                           #diagnostics.partnerConfig.sizeOfReceiveBuffer := 0;
                           #diagnostics.partnerConfig.sizeOfSendBuffer := 0;
                           #connected := #statConnected := TRUE;
                           #statState.cfgSender := #OPERATION;

                           #statDiag.bufferIndex := #statDiag.bufferIndex + 1;
                           #statDiag.buffer[#statDiag.bufferIndex].status := #STATUS_TCP_CONNECTED;
                           #statDiag.buffer[#statDiag.bufferIndex].subFunctionErrorID := 16#0000;
                           #statDiag.buffer[#statDiag.bufferIndex].additionalValue1 := 0.0;
                           #statDiag.buffer[#statDiag.bufferIndex].additionalValue2 := 0.0;
                           #statDiag.buffer[#statDiag.bufferIndex].additionalValue3 := 0.0;
                           #statDiag.buffer[#statDiag.bufferIndex].additionalValue4 := T#0ms;
                       END_IF;
                       //TCON still in progress
                   ELSE
                       IF (#diagnostics.localConfig.connection.isClient) THEN

                           #statDiag.bufferIndex := #statDiag.bufferIndex + 1;
                           #statDiag.buffer[#statDiag.bufferIndex].status := #STATUS_CLIENT_TRY_CONNECT;
                           #statDiag.buffer[#statDiag.bufferIndex].subFunctionErrorID := 16#0000;
                           #statDiag.buffer[#statDiag.bufferIndex].additionalValue1 := 0.0;
                           #statDiag.buffer[#statDiag.bufferIndex].additionalValue2 := 0.0;
                           #statDiag.buffer[#statDiag.bufferIndex].additionalValue3 := 0.0;
                           #statDiag.buffer[#statDiag.bufferIndex].additionalValue4 := T#0ms;
                       ELSE
                           #statDiag.bufferIndex := #statDiag.bufferIndex + 1;
                           #statDiag.buffer[#statDiag.bufferIndex].status := #STATUS_SERVER_PORT_OPEN;
                           #statDiag.buffer[#statDiag.bufferIndex].subFunctionErrorID := 16#0000;
                           #statDiag.buffer[#statDiag.bufferIndex].additionalValue1 := 0.0;
                           #statDiag.buffer[#statDiag.bufferIndex].additionalValue2 := 0.0;
                           #statDiag.buffer[#statDiag.bufferIndex].additionalValue3 := 0.0;
                           #statDiag.buffer[#statDiag.bufferIndex].additionalValue4 := T#0ms;
                       END_IF;
                   END_IF;
               END_REGION OPEN_CLIENT_SERVER

           #STATE_WAIT:
               REGION WAIT
                   //Wait and then establish the connection
                   IF (#statIterator > #STATE_WAIT) THEN

                       #tempConnOucId := 0;

                       //differ between different connection types (IPv4, QDN)
                       IF (#diagnostics.localConfig.connection.connectType = #CON_TYPE_IPV4) THEN
                           //IPv4
                           #instTCON(REQ := FALSE,
                                     ID := #statTconPar.ID,
                                     CONNECT := #statTconPar);
                           //store connection ID temporary
                           #tempConnOucId := #statTconPar.ID;
                       ELSE
                           //QDN (CON_TYPE_QDN)
                           #instTCON(REQ := FALSE,
                                     ID := #statTconParQdn.ID,
                                     CONNECT := #statTconParQdn);
                           //store connection ID temporary
                           #tempConnOucId := #statTconParQdn.ID;
                       END_IF;

                       #instTSEND(REQ := FALSE,
                                  ID := #tempConnOucId,
                                  DATA := #statSend.tsendFct.data);

                       #instTRCV(EN_R := FALSE,
                                 ID := #tempConnOucId,
                                 DATA := #statReceive.trcvFct.data);

                       #instTDISCON(REQ := FALSE,
                                    ID := #tempConnOucId);

                       IF (#diagnostics.localConfig.connection.isClient) THEN
                           #statState.connection := #OPEN_CLIENT;
                           #statTconPar.ActiveEstablished := TRUE;
                           #statTconParQdn.ActiveEstablished := TRUE;
                       ELSE
                           #statState.connection := #OPEN_SERVER;
                           #statTconPar.ActiveEstablished := FALSE;
                           #statTconParQdn.ActiveEstablished := FALSE;
                       END_IF;

                   ELSE
                       #statIterator := #statIterator + 1;
                   END_IF;
               END_REGION WAIT

           #FINISH_TSEND:
               REGION FINISH_TSEND
                   IF (#statIterator > #STATE_WAIT) THEN
                       #statIterator := 0;
                       #statState.connection := #FINISH_TRCV;
                   ELSE
                       //differ between different connection types (IPv4, QDN)
                       IF (#diagnostics.localConfig.connection.connectType = #CON_TYPE_IPV4) THEN
                           #tempConnOucId := #statTconPar.ID;
                       ELSE    //CON_TYPE_QDN
                           #tempConnOucId := #statTconParQdn.ID;
                       END_IF;

                       #instTSEND(REQ := TRUE,
                                  LEN := #statSend.tsendFct.dataOffset,
                                  ID := #tempConnOucId,
                                  DATA := #statSend.tsendFct.data,
                                  STATUS => #statSend.tsendFct.status);

                       IF ((#statSend.tsendFct.status = 16#0000) OR (#instTSEND.ERROR)) THEN
                           //"TSEND" instruction is finished
                           #statState.connection := #FINISH_TRCV;
                       ELSE
                           ;//"TSEND" instruction still in process
                       END_IF;
                   END_IF;
                   #statIterator := #statIterator + 1;
               END_REGION FINISH_TSEND

           #FINISH_TRCV:
               REGION FINISH_TRCV

                   IF (#statIterator > #STATE_WAIT) THEN
                       #statState.connection := #CALL_TDISCON;
                   ELSE
                       //differ between different connection types (IPv4, QDN)
                       IF (#diagnostics.localConfig.connection.connectType = #CON_TYPE_IPV4) THEN
                           #tempConnOucId := #statTconPar.ID;
                       ELSE    //CON_TYPE_QDN
                           #tempConnOucId := #statTconParQdn.ID;
                       END_IF;

                       #instTRCV(EN_R := TRUE,
                                 ID := #tempConnOucId,
                                 LEN := 0,
                                 ADHOC := TRUE,
                                 NDR => #statReceive.trcvFct.dataReceived,
                                 RCVD_LEN => #statReceive.trcvFct.dataLength,
                                 DATA := #statReceive.trcvFct.data);

                       //Is the "TRCV" instruction still in process
                       IF (#instTRCV.ERROR OR NOT #instTRCV.BUSY) THEN
                           #statState.connection := #CALL_TDISCON;
                       ELSE
                           ;//TRCV instruction still in process
                       END_IF;
                   END_IF;
                   #statIterator := #statIterator + 1;
               END_REGION FINISH_TRCV

           #CLOSE_CONNECTION:
               REGION CLOSE_CONNECTION
                   //reset FB Outputs
                   #connected := #statConnected := FALSE;
                   #sending := #statSending := FALSE;
                   #receivedDataLength := 0;
                   #error := FALSE;

                   //Is "TSEND" instruction still in process ?
                   IF (#statSend.tsendFct.status <> 16#0000) THEN
                       //"TSEND" instruction still in process
                       #statState.connection := #FINISH_TSEND;
                       #statIterator := 0;
                   ELSE
                       ;//"TSEND" instruction is finished
                   END_IF;

                   #instTRCV(EN_R := TRUE,
                             ID := #diagnostics.localConfig.connection.connectionID,
                             LEN := 0,
                             ADHOC := TRUE,
                             NDR => #statReceive.trcvFct.dataReceived,
                             RCVD_LEN => #statReceive.trcvFct.dataLength,
                             DATA := #statReceive.trcvFct.data);

                   //Is the "TRCV" instruction still in process
                   IF (#instTRCV.ERROR OR NOT #instTRCV.BUSY) THEN
                       #statState.connection := #CALL_TDISCON;
                   ELSE
                       #statState.connection := #FINISH_TRCV;
                       #statIterator := 0;
                   END_IF;
               END_REGION CLOSE_CONNECTION

           #CALL_TDISCON:
               REGION CALL_TDISCON
                   //differ between different connection types (IPv4, QDN)
                   IF (#diagnostics.localConfig.connection.connectType = #CON_TYPE_IPV4) THEN
                       #tempConnOucId := #statTconPar.ID;
                   ELSE    //CON_TYPE_QDN
                       #tempConnOucId := #statTconParQdn.ID;
                   END_IF;

                   #instTSEND(REQ := FALSE,
                              LEN := #statSend.tsendFct.dataOffset,
                              ID := #tempConnOucId,
                              DATA := #statSend.tsendFct.data);

                   #instTRCV(EN_R := FALSE,
                             ID := #diagnostics.localConfig.connection.connectionID,
                             LEN := 0,
                             ADHOC := TRUE,
                             NDR => #statReceive.trcvFct.dataReceived,
                             RCVD_LEN => #statReceive.trcvFct.dataLength,
                             DATA := #statReceive.trcvFct.data);

                   #instTDISCON(REQ := TRUE,
                                ID := #tempConnOucId);

                   //Error occurred during processing
                   IF (#instTDISCON.ERROR) THEN

                       #statDiag.bufferIndex := #statDiag.bufferIndex + 1;
                       #statDiag.buffer[#statDiag.bufferIndex].status := #ERR_CLOSE_CONNECTION;
                       #statDiag.buffer[#statDiag.bufferIndex].subFunctionErrorID := #instTDISCON.STATUS;
                       #statDiag.buffer[#statDiag.bufferIndex].additionalValue1 := 0.0;
                       #statDiag.buffer[#statDiag.bufferIndex].additionalValue2 := 0.0;
                       #statDiag.buffer[#statDiag.bufferIndex].additionalValue3 := 0.0;
                       #statDiag.buffer[#statDiag.bufferIndex].additionalValue4 := T#0ms;

                       #statState.connection := #STATE_INACTIVE_PREPARE;

                       #instTDISCON(REQ := FALSE,
                                    ID := #tempConnOucId);

                   ELSIF (#instTDISCON.DONE) THEN

                       #instTDISCON(REQ := FALSE,
                                    ID := #tempConnOucId);
                       //Job executed without errors
                       IF (#enable AND (NOT #statFallingEdgeEnable)) THEN
                           //Reconnect automatically if not in disconnecting process
                           #statIterator := 0;
                           #statState.connection := #STATE_WAIT;
                       ELSE
                           //Reset all active failures in the diagnostics buffer
                           FOR #statIterator := 0 TO #DIAG_BUFFER_UPPER_LIM BY 1 DO
                               #diagnostics.buffer[#statIterator].isActive := FALSE;
                           END_FOR;

                           #statState.connection := #STATE_INACTIVE_PREPARE;
                       END_IF;
                       //Job is not completed yet
                   ELSE
                       ;//Wait until job is finished
                   END_IF;
               END_REGION CALL_TDISCON

           #ERROR_STATE:
               REGION ERROR
                   ;
               END_REGION ERROR
       END_CASE;
   END_REGION STATE_MACHINE

   REGION DIAGNOSTICS
       // -----------------------------------------------------------------------------------------------------------
       //Diagnostics buffer
       // -----------------------------------------------------------------------------------------------------------
   diag:
       //Diagnostics entry is in the temp. buffer
       IF (#statDiag.bufferIndex <> -1) THEN

           //Get current time
           #statRet := RD_LOC_T(#tempActTime);
           //init
           #statDiag.actualIndex := 0;

           WHILE (#statDiag.actualIndex <= #statDiag.bufferIndex) DO

               #tempUDint := 0;
               //Check if the failure is already in the buffer and still active
               FOR #statIterator := 0 TO #DIAG_BUFFER_UPPER_LIM BY 1 DO

                   IF (#diagnostics.buffer[#statIterator].isActive = TRUE) THEN

                       IF ((#statDiag.buffer[#statDiag.actualIndex].status = #WARN_SEND_CYCLE_EXPIRED)
                           AND
                           (#diagnostics.buffer[#statIterator].status = #WARN_SEND_CYCLE_EXPIRED)
                           AND
                           (#diagnostics.buffer[#statIterator].additionalValue1 = #statDiag.buffer[#statDiag.actualIndex].additionalValue1)
                           AND
                           (#diagnostics.buffer[#statIterator].additionalValue2 = #statDiag.buffer[#statDiag.actualIndex].additionalValue2)
                           AND
                           (#diagnostics.buffer[#statIterator].additionalValue3 = #statDiag.buffer[#statDiag.actualIndex].additionalValue3)) THEN
                           //Retrigger just the activation time
                           #diagnostics.buffer[#statIterator].timestamp := #tempActTime;
                           #diagnostics.buffer[#statIterator].additionalValue4 := #statDiag.buffer[#statDiag.actualIndex].additionalValue4;
                           #tempUDint := 100;
                           EXIT;
                       ELSIF ((#diagnostics.buffer[#statIterator].status = #statDiag.buffer[#statDiag.actualIndex].status)
                           AND
                           (#diagnostics.buffer[#statIterator].additionalValue1 = #statDiag.buffer[#statDiag.actualIndex].additionalValue1)
                           AND
                           (#diagnostics.buffer[#statIterator].additionalValue2 = #statDiag.buffer[#statDiag.actualIndex].additionalValue2)
                           AND
                           (#diagnostics.buffer[#statIterator].additionalValue3 = #statDiag.buffer[#statDiag.actualIndex].additionalValue3)
                           AND
                           (#diagnostics.buffer[#statIterator].additionalValue4 = #statDiag.buffer[#statDiag.actualIndex].additionalValue4)) THEN
                           //Retrigger just the activation time
                           #diagnostics.buffer[#statIterator].timestamp := #tempActTime;
                           #tempUDint := 100;
                           EXIT;
                       ELSE
                           ;//ErrorId is not in the diagnostics buffer
                       END_IF;
                   END_IF;
               END_FOR;

               IF (#tempUDint = 100) THEN
                   ;//ErrorId was already retriggered
               ELSE
                   //Check range of diagnostics ring buffer [0...DIAG_ARRAY]
                   IF ((#diagnostics.bufferIndex = 255) OR (#diagnostics.bufferIndex = #DIAG_BUFFER_UPPER_LIM)) THEN
                       #diagnostics.bufferIndex := 0;
                   ELSE
                       #diagnostics.bufferIndex := #diagnostics.bufferIndex + 1;
                   END_IF;

                   //Stored new entry in the diagnostics buffer
                   #diagnostics.buffer[#diagnostics.bufferIndex].status := #statDiag.buffer[#statDiag.actualIndex].status;
                   #diagnostics.buffer[#diagnostics.bufferIndex].timestamp := #tempActTime;
                   #diagnostics.buffer[#diagnostics.bufferIndex].isActive := TRUE;

                   #diagnostics.buffer[#diagnostics.bufferIndex].subFunctionErrorID := #statDiag.buffer[#statDiag.actualIndex].subFunctionErrorID;
                   #diagnostics.buffer[#diagnostics.bufferIndex].additionalValue1 := #statDiag.buffer[#statDiag.actualIndex].additionalValue1;
                   #diagnostics.buffer[#diagnostics.bufferIndex].additionalValue2 := #statDiag.buffer[#statDiag.actualIndex].additionalValue2;
                   #diagnostics.buffer[#diagnostics.bufferIndex].additionalValue3 := #statDiag.buffer[#statDiag.actualIndex].additionalValue3;
                   #diagnostics.buffer[#diagnostics.bufferIndex].additionalValue4 := #statDiag.buffer[#statDiag.actualIndex].additionalValue4;
               END_IF;

               IF ((#diagnostics.buffer[#diagnostics.bufferIndex].status = #STATUS_TCP_CONNECTED)
                   OR (#diagnostics.buffer[#diagnostics.bufferIndex].status = #STATUS_CONNECTED_V1)
                   OR (#diagnostics.buffer[#diagnostics.bufferIndex].status = #STATUS_CONNECTED_V2))
               THEN
                   #statConnectAttempts := 0;
                   #diagnostics.statistics.lastConnect := #tempActTime;
               END_IF;

               //Set FB status
               #status := #statStatus := #statDiag.buffer[#statDiag.actualIndex].status;

               //Check if FB.error has been set ?
               IF ((#statDiag.buffer[#statDiag.actualIndex].status >= #ERR_COM_SERVICE)//16#8200
                   AND
                   (#statDiag.buffer[#statDiag.actualIndex].status <= #ERR_WRONG_TELEGRAM_ID))//16#8614
               THEN

                   #error := TRUE;
                   #connected := #statConnected := FALSE;
                   #sending := #statSending := FALSE;
                   #dataReceived := #statDataReceived := FALSE;
                   #receivedDataLength := 0;

                   //Check if FB.busy has been set ?
                   IF ((#statDiag.buffer[#statDiag.actualIndex].status >= #ERR_OPEN_CLIENT)//16#8600
                       AND
                       (#statDiag.buffer[#statDiag.actualIndex].status <= #ERR_WRONG_TELEGRAM_ID))//16#8614
                   THEN
                       #busy := TRUE;
                   ELSE
                       #busy := FALSE;
                   END_IF;

                   EXIT;//Leave loop
               ELSE
                   ;
               END_IF;

               //Increase index
               #statDiag.actualIndex := #statDiag.actualIndex + 1;

           END_WHILE;
       ELSE
           ;//No failure
       END_IF;//End: Diagnostics buffer
   END_REGION DIAGNOSTICS
END_FUNCTION_BLOCK

FUNCTION_BLOCK "GateAccess_Station_FB"   // FB26, SCL
{ S7_Optimized_Access := 'TRUE' }
VERSION : 0.1
// stored: AutoNumber true, IsIECCheckEnabled false, IsRetainMemResEnabled false, MemoryReserve 100, SetENOAutomatically false, UDAEnableTagReadback false
   VAR_INPUT
      Sys_No : UInt;
      Right_True { ExternalAccessible := 'False'; ExternalVisible := 'False'; ExternalWritable := 'False'} : Bool;
      Switches { ExternalAccessible := 'False'; ExternalVisible := 'False'; ExternalWritable := 'False'} : Byte;
      GateLockedFeedback : Bool;
      NoEStop : Bool;
      I_G1_GuardOpen : Bool;
      I_L1_Unlocked : Bool;
      FaultResetCmd : Bool;
      AllDrivesHealthy : Bool;
      SafetyResetDone : Bool;
      NoVTDLocalMode : Bool;
      NoCrossoverPaused : Bool;
      Safe_Bypassed : Bool;
      LGX_Secure_Access : Bool;
      AllDevicesStopped : Bool;
   END_VAR
   VAR_OUTPUT
      Lamps { ExternalAccessible := 'False'; ExternalVisible := 'False'; ExternalWritable := 'False'} : Byte;
      O_S1_SolenoidEnergise : Bool;
      "Lock Reset" { ExternalAccessible := 'False'; ExternalVisible := 'False'; ExternalWritable := 'False'} : Bool;
      CurrentState : UInt;
      GateFault : Bool;
   END_VAR
   VAR_IN_OUT
      Gate_Station : "Gate_Station_UDT";
   END_VAR
   VAR
      RTE_PB : Bool;
      Reset_PB : Bool;
      Restart_PB : Bool;
      GateAccessControl : "GateAccessControl_FB";
      ModeManager : "ModeManager_FB";
   END_VAR
   VAR_TEMP
      i : UInt;
   END_VAR
   VAR CONSTANT
      AUTO_RUNNING : UInt := 0;
      RTE_REQUESTED : UInt := 1;
      SAFE_TO_UNLOCK : UInt := 3;
      ACCESS_MANUAL_MODE : UInt := 4;
      RESETTING : UInt := 6;
   END_VAR
BEGIN
   // IF #Right_True THEN
   //     // #Switches
   //     #Reset_PB := #Switches.%X1; //Blue button - Restart_PB
   //     #Restart_PB := #Switches.%X2; //White button - Reset_PB
   //     #RTE_PB := #Switches.%X3; //Green button - RTE_PB
   // ELSE
   // //     //Switches
   //     #Restart_PB := #Switches.%X1; //White button - Reset_PB
   //     #Reset_PB := #Switches.%X2; //Blue button - Restart_PB
   //     #RTE_PB := #Switches.%X3; //Green button - RTE_PB
   // END_IF;
   IF #Right_True THEN
       // #Switches
       #Reset_PB := #Switches.%X1; //Blue button - Reset_PB
       #Restart_PB := #Switches.%X3; //Green button - Restart_PB
       #RTE_PB := #Switches.%X2; //White button - RTE_PB
   ELSE
       //Switches
       #Restart_PB := #Switches.%X3; //Green button - Restart_PB
       #Reset_PB := #Switches.%X2; //Blue button - Reset_PB
       #RTE_PB := #Switches.%X1; //White button - RTE_PB
   END_IF;

   // ------------------------------------------------------
   // Step 1: run the hardware interface FB, feeding it the
   // consolidated safety signals read directly from
   // DB_SafetyLogic for this gate. GateClosed and
   // ForceRTE_Request come out ready for ModeManager below.
   // ------------------------------------------------------
   #GateAccessControl(
                      UnlockPermissive := #ModeManager.GateUnlockPermissive,
                      FaultResetCmd := #FaultResetCmd,
                      I_G1_GuardOpen := #I_G1_GuardOpen,
                      I_L1_Unlocked := #I_L1_Unlocked,
                      GateLockedFeedback := #GateLockedFeedback,
                      NoEStop := #NoEStop
   );

   // ------------------------------------------------------
   // Step 2: run the mode state machine, feeding it the
   // fresh feedback from GateAccessControl plus the same
   // consolidated safety signals and cross-subsystem
   // interlocks.
   // ------------------------------------------------------
   #ModeManager(
                RTE_PB := #RTE_PB,
                Reset_PB := #Reset_PB,
                Restart_PB := #Restart_PB,
                GateClosed := #GateAccessControl.GateClosed,
                GateLockedFeedback := #GateLockedFeedback,
                GateFault := #GateAccessControl.GateFault,
                NoEStop := #NoEStop,
                AllDrivesHealthy := #AllDrivesHealthy,
                SafetyResetDone := #SafetyResetDone,
                NoVTDLocalMode := #NoVTDLocalMode,
                NoCrossoverPaused := #NoCrossoverPaused,
                AllDevicesStopped := #Gate_Station.Secure_Access AND #AllDevicesStopped AND #LGX_Secure_Access,
                Safe_Bypassed := #Safe_Bypassed,
                ForceRTE := #GateAccessControl.ForceRTE_Request,
                Reset := #FaultResetCmd
   );

   // ------------------------------------------------------
   // Step 3: expose local outputs for the physical wiring.
   // ------------------------------------------------------
   #O_S1_SolenoidEnergise := #GateAccessControl.O_S1_SolenoidEnergise;
   #CurrentState := #ModeManager.CurrentState;
   #GateFault := #GateAccessControl.GateFault;

   //Send all devices to automatic mode
   IF #ModeManager.CurrentState = #RESETTING AND #Sys_No <> 0 THEN
       FOR #i := "Settings_DB".VTD_Sys[#Sys_No].Lowest_Level TO "Settings_DB".VTD_Sys[#Sys_No].Highest_Level DO
           "Control_DB".VTD_Sys[#Sys_No].Instruction.Reset :=
           "Control_DB".ECnv_Sys[#Sys_No].Instruction.Reset :=
           "Control_DB".LCnv_Sys[#Sys_No].Cnv_Level[#i].Cnv1.Instruction.Reset :=
           "Control_DB".LCnv_Sys[#Sys_No].Cnv_Level[#i].Cnv2.Instruction.Reset := TRUE;
       END_FOR;

       IF #AllDrivesHealthy THEN
           FOR #i := "Settings_DB".VTD_Sys[#Sys_No].Lowest_Level TO "Settings_DB".VTD_Sys[#Sys_No].Highest_Level DO
               "Control_DB".VTD_Sys[#Sys_No].Instruction.Reset :=
               "Control_DB".ECnv_Sys[#Sys_No].Instruction.Reset :=
               "Control_DB".LCnv_Sys[#Sys_No].Cnv_Level[#i].Cnv1.Instruction.Reset :=
               "Control_DB".LCnv_Sys[#Sys_No].Cnv_Level[#i].Cnv2.Instruction.Reset := FALSE;
           END_FOR;

           FOR #i := "Settings_DB".VTD_Sys[#Sys_No].Lowest_Level TO "Settings_DB".VTD_Sys[#Sys_No].Highest_Level DO
               "Control_DB".VTD_Sys[#Sys_No].Instruction.Mode_Change :=
               "Control_DB".ECnv_Sys[#Sys_No].Instruction.Mode_Change :=
               "Control_DB".LCnv_Sys[#Sys_No].Cnv_Level[#i].Cnv1.Instruction.Mode_Change :=
               "Control_DB".LCnv_Sys[#Sys_No].Cnv_Level[#i].Cnv2.Instruction.Mode_Change :=
               "Control_DB".LCnv_Sys[#Sys_No].Cnv_Level[#i].Cnv1.Safety_Stop_Cnrl.Mode :=
               "Control_DB".LCnv_Sys[#Sys_No].Cnv_Level[#i].Cnv2.Safety_Stop_Cnrl.Mode := 3;

               "Control_DB".VTD_Sys[#Sys_No].Instruction.Enable :=
               "Control_DB".ECnv_Sys[#Sys_No].Instruction.Enable :=
               "Control_DB".LCnv_Sys[#Sys_No].Cnv_Level[#i].Cnv1.Instruction.Enable :=
               "Control_DB".LCnv_Sys[#Sys_No].Cnv_Level[#i].Cnv2.Instruction.Enable := TRUE;
           END_FOR;
       END_IF;
   END_IF;

   //Send all devices to manual mode
   IF #ModeManager.CurrentState = #ACCESS_MANUAL_MODE AND #Sys_No <> 0 THEN
       FOR #i := "Settings_DB".VTD_Sys[#Sys_No].Lowest_Level TO "Settings_DB".VTD_Sys[#Sys_No].Highest_Level DO
           "Control_DB".VTD_Sys[#Sys_No].Instruction.Mode_Change :=
           "Control_DB".ECnv_Sys[#Sys_No].Instruction.Mode_Change :=
           "Control_DB".LCnv_Sys[#Sys_No].Cnv_Level[#i].Cnv1.Instruction.Mode_Change :=
           "Control_DB".LCnv_Sys[#Sys_No].Cnv_Level[#i].Cnv2.Instruction.Mode_Change :=
           "Control_DB".LCnv_Sys[#Sys_No].Cnv_Level[#i].Cnv1.Safety_Stop_Cnrl.Mode :=
           "Control_DB".LCnv_Sys[#Sys_No].Cnv_Level[#i].Cnv2.Safety_Stop_Cnrl.Mode := 1;
       END_FOR;
   END_IF;

   // IF #Right_True THEN
   //     #Lamps.%X0 := (NOT #NoEStop OR #GateAccessControl.GateFault) AND "Clock_1Hz"; //Estop lamp
   //     #Lamps.%X2 := #ModeManager.ReqFlash_RestartLamp AND "Clock_1Hz"; //White lamp - Restart_PB
   //     #Lamps.%X1 := #ModeManager.ReqFlash_ResetLamp AND "Clock_1Hz"; //Blue lamp - Reset_PB
   //     #Lamps.%X3 := #ModeManager.RestartLampSteadyOn OR #ModeManager.ReqFlash_RTE_Lamp; //Green lamp - RTE_PB
   // ELSE
   //     #Lamps.%X0 := (NOT #NoEStop OR #GateAccessControl.GateFault) AND "Clock_1Hz"; //Estop lamp
   //     #Lamps.%X2 := #ModeManager.ReqFlash_ResetLamp  AND "Clock_1Hz"; //Blue lamp - Reset_PB
   //     #Lamps.%X1 := #ModeManager.ReqFlash_RestartLamp AND "Clock_1Hz"; //White lamp - Restart_PB
   //     #Lamps.%X3 := #ModeManager.RestartLampSteadyOn OR #ModeManager.ReqFlash_RTE_Lamp; //Green lamp - RTE_PB
   // END_IF;
   IF #Right_True THEN
       #Lamps.%X0 := (NOT #NoEStop OR #GateAccessControl.GateFault) AND "Clock_1Hz"; //Estop lamp
       #Lamps.%X3 := (#ModeManager.ReqFlash_RestartLamp AND "Clock_1Hz") OR #ModeManager.RestartLampSteadyOn; //Green lamp - Restart_PB
       #Lamps.%X1 := #ModeManager.ReqFlash_ResetLamp AND "Clock_1Hz"; //Blue lamp - Reset_PB
       #Lamps.%X2 := #ModeManager.ReqFlash_RTE_Lamp OR (#ModeManager.CurrentState = #SAFE_TO_UNLOCK AND NOT #NoEStop) OR #ModeManager.CurrentState = #SAFE_TO_UNLOCK OR #ModeManager.CurrentState = #ACCESS_MANUAL_MODE; //White lamp - RTE_PB
   ELSE
       #Lamps.%X0 := (NOT #NoEStop OR #GateAccessControl.GateFault) AND "Clock_1Hz"; //Estop lamp
       #Lamps.%X2 := #ModeManager.ReqFlash_ResetLamp AND "Clock_1Hz"; //Blue lamp - Reset_PB
       #Lamps.%X3 := (#ModeManager.ReqFlash_RestartLamp AND "Clock_1Hz") OR #ModeManager.RestartLampSteadyOn; //Green lamp - Restart_PB
       #Lamps.%X1 := #ModeManager.ReqFlash_RTE_Lamp OR (#ModeManager.CurrentState = #SAFE_TO_UNLOCK AND NOT #NoEStop) OR #ModeManager.CurrentState = #SAFE_TO_UNLOCK OR #ModeManager.CurrentState = #ACCESS_MANUAL_MODE; //White lamp - RTE_PB
   END_IF;

   //Gate station control
   //
   #Gate_Station.Requested_Access := #ModeManager.CurrentState = #RTE_REQUESTED;
   #Gate_Station.Safe_To_Restart := #ModeManager.RestartLampSteadyOn;
END_FUNCTION_BLOCK

FUNCTION_BLOCK "GateAccessControl_FB"   // FB23, SCL
{ S7_Optimized_Access := 'TRUE' }
VERSION : 0.1
// stored: AutoNumber true, IsIECCheckEnabled false, IsRetainMemResEnabled false, MemoryReserve 100, SetENOAutomatically false, UDAEnableTagReadback false
   VAR_INPUT
      UnlockPermissive : Bool;   // TRUE = ModeManager allows gate to be unlocked
      FaultResetCmd : Bool;   // rising edge = attempt to reset a latched GateFault (only if hardware is OK)
      I_G1_GuardOpen : Bool;   // BYTE1 bit0: Guard Open(1) / Guard Closed(0)
      I_L1_Unlocked : Bool;   // BYTE2 bit0: Unlocked(1) / Locked(0) - diagnostic only, NOT safety-relevant
      GateLockedFeedback : Bool;   // Guard switch safe output. Closed+Locked=1
      NoEStop : Bool;   // E-Stop safe output. Released=1
      ResetPulseTime : Time := T#500MS;   // R1 / RS_xx pulse width
      LockConfirmTimeout : Time := T#300S;   // max time allowed for lock feedback to confirm after command
      UnlockConfirmTimeout : Time := T#300S;   // max time allowed for unlock feedback to confirm after command
   END_VAR
   VAR_OUTPUT
      O_S1_SolenoidEnergise : Bool;   // BYTE1 bit0: Energise(1) / De-energise(0) // ASSUMPTION: Energise = UNLOCK (fail-safe locked // when de-energised). CONFIRM against your GSDML / // wiring before commissioning - if reversed, invert // the assignment below.
      GateClosed : Bool;   // debounced gate closed status
      GateFault : Bool;   // latched TRUE on lock/unlock discrepancy timeout
      ForceRTE_Request : Bool;   // pulses TRUE to force ModeManager into RTE_REQUESTED // (e.g. rear escape used unexpectedly - area accessed // outside the normal sequence, treat as if entry // was requested so the system re-syncs its state)
   END_VAR
   VAR
      ResetPulse_GuardReset { S7_SetPoint := 'True'} : TP_TIME;
      LockConfirmTON { S7_SetPoint := 'True'} : TON_TIME;
      UnlockConfirmTON { S7_SetPoint := 'True'} : TON_TIME;
      FaultResetCmd_Edge_M { S7_SetPoint := 'True'} : Bool;
      FaultResetCmd_Rising : Bool;
      GateFault_Latch : Bool;
      WasLockedAndValid : Bool;
   END_VAR
BEGIN
   // ------------------------------------------------------
   // Standard feedback passthrough
   // ------------------------------------------------------
   #GateClosed := NOT #I_G1_GuardOpen;

   // ------------------------------------------------------
   // Solenoid command.
   // Energise = Unlock, confirmed by user: solenoid energised
   // frees the mechanism so the operator can rotate the manual
   // handle. De-energised = locked (fail-safe default).
   // ------------------------------------------------------
   #O_S1_SolenoidEnergise := #UnlockPermissive AND NOT #GateFault_Latch;

   // ------------------------------------------------------
   // Lock / unlock confirmation supervision, using the
   // consolidated GateLockedFeedback signal fed in from the
   // safety logic.
   // ------------------------------------------------------
   #LockConfirmTON(IN := NOT #O_S1_SolenoidEnergise AND NOT #GateLockedFeedback AND #GateClosed,
                   PT := #LockConfirmTimeout);
   IF #LockConfirmTON.Q THEN
       (*#GateFault_Latch := TRUE*);
   END_IF;

   #UnlockConfirmTON(IN := #O_S1_SolenoidEnergise AND #GateLockedFeedback,
                     PT := #UnlockConfirmTimeout);
   IF #UnlockConfirmTON.Q THEN
       (*#GateFault_Latch := TRUE*);
   END_IF;

   // ------------------------------------------------------
   // Forced-open / unexpected drop detection.
   // If the gate was locked last scan and is no longer locked
   // THIS scan, without an unlock having been permitted, this
   // mirrors the device's own "Guard forced open, reset
   // required" condition (LS red double flash).
   // ------------------------------------------------------
   IF #WasLockedAndValid AND NOT #GateLockedFeedback AND NOT #UnlockPermissive THEN
       // #GateFault_Latch := TRUE;
       (*#ForceRTE_Request := TRUE*);
   ELSE
       #ForceRTE_Request := FALSE;
   END_IF;

   #WasLockedAndValid := #GateLockedFeedback;

   // ------------------------------------------------------
   // Reset sequence: pulse R1 (guard reset), per manual
   // procedure. Safe qualifier resets (RS_GSx/RS_ESx) are
   // now the responsibility of the separate safety logic
   // block, not this one.
   // ------------------------------------------------------
   #FaultResetCmd_Rising := #FaultResetCmd AND NOT #FaultResetCmd_Edge_M;
   #FaultResetCmd_Edge_M := #FaultResetCmd;

   #ResetPulse_GuardReset(IN := #FaultResetCmd_Rising,
                          PT := #ResetPulseTime);

   IF #FaultResetCmd_Rising
       AND NOT #LockConfirmTON.Q
       AND NOT #UnlockConfirmTON.Q
       AND #GateClosed THEN
       #GateFault_Latch := FALSE;
   END_IF;

   #GateFault := #GateFault_Latch := FALSE;
END_FUNCTION_BLOCK

FUNCTION_BLOCK "ModeManager_FB"   // FB8, SCL
{ S7_Optimized_Access := 'TRUE' }
VERSION : 0.1
// stored: AutoNumber true, IsIECCheckEnabled false, IsRetainMemResEnabled false, MemoryReserve 100, SetENOAutomatically false, UDAEnableTagReadback false
   VAR_INPUT
      RTE_PB : Bool;   // Request To Enter pushbutton, rising edge triggers request
      Reset_PB : Bool;   // Reset pushbutton, rising edge triggers reset attempt
      Restart_PB : Bool;   // Restart pushbutton, rising edge triggers return to auto
      ForceRTE : Bool;   // one-scan pulse from FB_GateAccessControl.ForceRTE_Request
      GateClosed : Bool;   // TRUE = gate physically closed
      GateLockedFeedback : Bool;   // TRUE = gate lock solenoid confirmed locked
      GateFault : Bool;   // from FB_GateAccessControl - blocks Auto/Restart
      NoEStop : Bool;   // TRUE = no emergency stop active anywhere in chain
      AllDrivesHealthy : Bool;   // TRUE = no drive faults on VTD/shuttle drives
      SafetyResetDone : Bool;   // TRUE = upstream safety reset permissive satisfied
      NoVTDLocalMode : Bool;   // TRUE = no VTD station currently in Local mode
      NoCrossoverPaused : Bool;   // TRUE = no conveyor crossover currently paused
      AllDevicesStopped : Bool;   // TRUE = all VTDs confirmed at standstill
      Safe_Bypassed : Bool;
      Reset : Bool;
   END_VAR
   VAR_OUTPUT
      CurrentState : UInt;   // current sequence state, for HMI/diagnostics
      GateUnlockPermissive : Bool;   // TRUE = safe to unlock gate solenoid (SAFE_TO_UNLOCK onwards)
      StopNewAutoCycles : Bool;   // TRUE = do not start new automatic cycles
      AutoModeAllowed : Bool;   // TRUE = auto mode is permitted (all interlocks satisfied)
      ManualModeActive : Bool;   // TRUE = system is in manual/jog/local maintenance mode
      ReqFlash_RTE_Lamp : Bool;
      ReqFlash_ResetLamp : Bool;
      ReqFlash_RestartLamp : Bool;
      RestartLampSteadyOn : Bool;
      RTE_LampSteadyOn : Bool;
   END_VAR
   VAR
      RTE_PB_Rising : Bool;   // edge memory for RTE_PB
      Reset_PB_Rising : Bool;   // edge memory for Reset_PB
      Restart_PB_Rising : Bool;   // edge memory for Restart_PB
      T_Delay_DB { S7_SetPoint := 'True'} : TON_TIME;
      EStop_Pressed : Bool;
      PLCInitialization : Bool;
   END_VAR
   VAR_TEMP
      RTE_PB_Edge_M : Bool;   // temp for R_TRIG-style edge detection
      Reset_PB_Edge_M : Bool;
      Restart_PB_Edge_M : Bool;
   END_VAR
   VAR CONSTANT
      AUTO_RUNNING : UInt := 0;
      RTE_REQUESTED : UInt := 1;
      SAFE_BYPASS : UInt := 2;
      SAFE_TO_UNLOCK : UInt := 3;
      ACCESS_MANUAL_MODE : UInt := 4;
      READY_TO_RESET : UInt := 5;
      RESETTING : UInt := 6;
      READY_TO_RESTART : UInt := 7;
   END_VAR
BEGIN
   #RTE_PB_Rising := #RTE_PB AND NOT #RTE_PB_Edge_M;
   #Reset_PB_Rising := #Reset_PB AND NOT #Reset_PB_Edge_M;
   #Restart_PB_Rising := #Restart_PB AND NOT #Restart_PB_Edge_M;

   #RTE_PB_Edge_M := #RTE_PB;
   #Reset_PB_Edge_M := #Reset_PB;
   #Restart_PB_Edge_M := #Restart_PB;

   IF #Reset THEN
       #CurrentState := #AUTO_RUNNING;
   END_IF;

   // Emergency Access
   // 
   IF "FirstScan" THEN
       #PLCInitialization := TRUE;
   ELSIF "Reset_All" AND #NoEStop THEN
       #PLCInitialization := FALSE;
   END_IF;

   IF NOT #PLCInitialization THEN
       IF NOT #NoEStop AND NOT #EStop_Pressed THEN
           #CurrentState := #SAFE_TO_UNLOCK;
           #EStop_Pressed := TRUE;
       ELSIF #NoEStop THEN
           #EStop_Pressed := FALSE;
       END_IF;
   END_IF;

   CASE #CurrentState OF

       #AUTO_RUNNING:
           IF #RTE_PB_Rising THEN
               #CurrentState := #RTE_REQUESTED;
           END_IF;

       #RTE_REQUESTED:
           IF #AllDevicesStopped THEN
               #CurrentState := #SAFE_BYPASS;
           END_IF;

       #SAFE_BYPASS:
           IF #Safe_Bypassed THEN
               #T_Delay_DB(IN:=TRUE,
                           PT:=T#500MS);
               IF #T_Delay_DB.Q THEN
                   #T_Delay_DB(IN := FALSE,
                               PT := T#0MS);
                   #CurrentState := #SAFE_TO_UNLOCK;
               END_IF;
           END_IF;

       #SAFE_TO_UNLOCK:
           // Solenoid is now de-energised->energised per GateUnlockPermissive,
           // which physically frees the mechanism so the operator can rotate
           // the manual handle. Transition to manual mode once the gate is
           // actually opened.
           IF NOT #GateClosed THEN
               #CurrentState := #ACCESS_MANUAL_MODE;
           END_IF;

       #ACCESS_MANUAL_MODE:
           // Gate physically closed again (handle rotated back, solenoid
           // still energised/unlocked at this point - lock only re-engages
           // in RESETTING once Reset is pressed).
           IF #GateClosed THEN
               #CurrentState := #READY_TO_RESET;
           END_IF;

       #READY_TO_RESET:
           IF #Reset_PB_Rising THEN
               #CurrentState := #RESETTING;
           END_IF;

       #RESETTING:
           // Lock is commanded via GateUnlockPermissive=FALSE
           // (see output mapping below); wait for GS1/GS2 to
           // confirm locked before allowing restart readiness.
           IF #GateLockedFeedback AND #SafetyResetDone AND #NoVTDLocalMode AND NOT #GateFault AND #AllDrivesHealthy THEN
               #CurrentState := #READY_TO_RESTART;
           END_IF;

       #READY_TO_RESTART:
           IF #Restart_PB_Rising
               AND #NoEStop
               AND NOT #GateFault
               AND #AllDrivesHealthy
               AND #NoVTDLocalMode
               AND #NoCrossoverPaused THEN
               #CurrentState := #AUTO_RUNNING;
           END_IF;

   END_CASE;

   // ------------------------------------------------------
   // OUTPUT MAPPING
   // ------------------------------------------------------
   // GateUnlockPermissive drives O_S1_SolenoidEnergise (assumed
   // energise=unlock) in FB_GateAccessControl. In RESETTING /
   // READY_TO_RESTART / AUTO_RUNNING the gate must be LOCKED,
   // so permissive is FALSE (commands lock, per assumption).
   #GateUnlockPermissive := (#CurrentState = #SAFE_TO_UNLOCK)
   OR (#CurrentState = #ACCESS_MANUAL_MODE)
   // OR (#CurrentState = #READY_TO_RESET)
   ;

   #StopNewAutoCycles := NOT (#CurrentState = #AUTO_RUNNING);
   #ManualModeActive := (#CurrentState = #ACCESS_MANUAL_MODE);

   #AutoModeAllowed := (#CurrentState = #AUTO_RUNNING)
   AND #GateClosed
   AND #GateLockedFeedback
   AND #NoEStop
   AND NOT #GateFault
   // AND #NoVTDLocalMode
   AND #NoCrossoverPaused
   AND #AllDrivesHealthy
   AND #SafetyResetDone;

   #RestartLampSteadyOn := (#CurrentState = #AUTO_RUNNING);
   #RTE_LampSteadyOn := (#CurrentState = #SAFE_TO_UNLOCK);
   #ReqFlash_RTE_Lamp := (#CurrentState = #RTE_REQUESTED) AND "Clock_1Hz";
   #ReqFlash_ResetLamp := (#CurrentState = #READY_TO_RESET);
   #ReqFlash_RestartLamp := (#CurrentState = #READY_TO_RESTART);
END_FUNCTION_BLOCK

FUNCTION_BLOCK "Order_Table_FB"   // FB31, SCL
{ S7_Optimized_Access := 'TRUE' }
VERSION : 0.1
// stored: AutoNumber false, IsIECCheckEnabled false, IsRetainMemResEnabled false, MemoryReserve 100, SetENOAutomatically false, UDAEnableTagReadback false
   VAR_INPUT
      System_Selected { ExternalWritable := 'False'} : Bool;
      AutoMan_Switch : Bool;   // Auto/Man Switch on CPU Panel - 1 = Auto, 0 = Manual
      CurrentTime { ExternalWritable := 'False'} : String;
      CurrentDTL : DTL;
      Watchdog : "Watchdog_Settings_UDT";
      OPC_UA_State_VTD : UInt;
      OPC_UA_State_Shuttle : UInt;
      OPC_UA_State_CNV : UInt;
      Clear_OrderTable : Bool;
   END_VAR
   VAR_IN_OUT
      VTD : "VTD_Control";
      Extrator_Conveyor : "ECnv_Control";
      Cnv_Buffer_11 : "Buffer_Cnv_Control";
      Cnv_Buffer_21 : "Buffer_Cnv_Control";
      Cnv_Buffer_31 : "Buffer_Cnv_Control";
      Cnv_Buffer_41 : "Buffer_Cnv_Control";
      Cnv_Buffer_51 : "Buffer_Cnv_Control";
      Cnv_Buffer_61 : "Buffer_Cnv_Control";
      Cnv_Buffer_71 : "Buffer_Cnv_Control";
      Cnv_Buffer_81 : "Buffer_Cnv_Control";
      Cnv_Buffer_12 : "Buffer_Cnv_Control";
      Cnv_Buffer_22 : "Buffer_Cnv_Control";
      Cnv_Buffer_32 : "Buffer_Cnv_Control";
      Cnv_Buffer_42 : "Buffer_Cnv_Control";
      Cnv_Buffer_52 : "Buffer_Cnv_Control";
      Cnv_Buffer_62 : "Buffer_Cnv_Control";
      Cnv_Buffer_72 : "Buffer_Cnv_Control";
      Cnv_Buffer_82 : "Buffer_Cnv_Control";
      System : "System_UDT";
      Control_OPC_Ua : "WMS_OPC_UA";
   END_VAR
   VAR
      VTD_CurrentOrder { ExternalWritable := 'False'} : UDInt := 0;
      Pallet_InOut_CurrentOrder : UDInt;
      Shuttle_InOut_CurrentOrder : UDInt;
      VTDDoneRTrig : R_TRIG;
      Pallet_InOut_RTrig { S7_SetPoint := 'True'} : R_TRIG;
      Shuttle_InOut_RTrig { S7_SetPoint := 'True'} : R_TRIG;
      PalletRefused_RTrig { ExternalWritable := 'False'} : R_TRIG;
      ErrorRTrig { ExternalWritable := 'False'} : R_TRIG;
      CancelRTrig { ExternalWritable := 'False'} : R_TRIG;
      PauseRTrig { ExternalWritable := 'False'} : R_TRIG;
      ResumeRTrig { ExternalWritable := 'False'} : R_TRIG;
      Clear_Store : R_TRIG;
      Clear_Retrieve : R_TRIG;
      Canceling : Bool;
      VTD_WatchdogTimer : TON_TIME;
      Pallet_InOut_WatchdogTimer { S7_SetPoint := 'True'} : TON_TIME;
      Shuttle_InOut_WatchdogTimer { S7_SetPoint := 'True'} : TON_TIME;
      VTD_WatchdogStart : Bool;
      Pallet_InOut_WatchdogStart : Bool;
      Shuttle_InOut_WatchdogStart : Bool;
      F_AutoMode { S7_SetPoint := 'True'} : F_TRIG;
   END_VAR
   VAR_TEMP
      i : DInt;
      n : DInt;
      EmptyOrder : "OrderTable_UDT";
      MaxRunningOrderNo : UInt;
   END_VAR
   VAR CONSTANT
      VTD_DEVICE : String := 'VTD';
      PALLET_INOUT_DEVICE : String := 'Pallet In Out';
      SHUTTLE_INOUT_DEVICE : String := 'Shuttle In Out';
      RUNNING_STATUS : String := 'Running';
      COMPLETED_STATUS : String := 'Completed';
      QUEUED_STATUS : String := 'Queued';
      PALLET_REFUSED_STATUS : String := 'Pallet Refused';
      ERROR_STATUS : String := 'Error';
      CANCELED_STATUS : String := 'Canceled';
      PAUSED_STATUS : String := 'Paused';
      ORDER_REFUSED : String := 'Refused';
      ERROR_CANCELED_STATUS : String := 'Error\Cancel';
   END_VAR
BEGIN

   // Converts the task type for strings 
   IF #System.OrderTable[1].OPC_Control.Task_Type = 1 THEN
       #System.OrderTable[1].Device := 'VTD';
   ELSIF #System.OrderTable[1].OPC_Control.Task_Type = 4 OR #System.OrderTable[1].OPC_Control.Task_Type = 5  THEN
       #System.OrderTable[1].Device := 'Pallet In Out';
   ELSIF #System.OrderTable[1].OPC_Control.Task_Type = 2 OR #System.OrderTable[1].OPC_Control.Task_Type = 3 THEN
       #System.OrderTable[1].Device := 'Shuttle In Out';
   ELSE
       #System.OrderTable[1].Device := '';
   END_IF;

   REGION #New Order was Sent
       IF #System.OrderSent THEN
           //Count orders in Step Table
           FOR #i := 0 TO 20 DO
               IF #System.StepTable[#i].OrderNo <> 0
                   AND #System.StepTable[#i].StepNo <> 0
                   AND #System.StepTable[#i].PlaceTime <> ''
               THEN
                   #System.StepTable[#i].Status := #QUEUED_STATUS;
                   #n += 1;
               ELSE
                   EXIT;
               END_IF;
           END_FOR;
           IF #n > 0 THEN
               //shift order table down by Order number rows
               FOR #i := 99 TO (#n + 1) BY -1 DO
                   #System.OrderTable[#i] := #System.OrderTable[#i - #n];
               END_FOR;
               //copy data from step table to order table
               FOR #i := 0 (*1*) TO #n DO
                   #System.OrderTable[#n - #i (*+ 1*)] := #System.StepTable[#i];
               END_FOR;
               //clean step table
               FOR #i := 0 (*1*) TO 20 DO
                   #System.StepTable[#i] := #EmptyOrder;
               END_FOR;
               #System.CurrentOrder += #n;

               //VTD move to floor
               IF #VTD_CurrentOrder <> 0 THEN
                   #VTD_CurrentOrder += #n;
               END_IF;

               //Shuttle transfer in/out of the VTD
               IF #Pallet_InOut_CurrentOrder <> 0 THEN
                   #Pallet_InOut_CurrentOrder += #n;
               END_IF;

               //Shuttle in/out of the VTD
               IF #Shuttle_InOut_CurrentOrder <> 0 THEN
                   #Shuttle_InOut_CurrentOrder += #n;
               END_IF;

                       END_IF;
           #System.OrderSent := FALSE;
       END_IF;
   END_REGION

   REGION Auto/Man Mode
       //Enable Devices in Auto/Man Mode
       IF #System.Auto_Man THEN
           // #VTD.Mode := #Extrator_Conveyor.Mode := #Cnv_Buffer_1.Mode := #Cnv_Buffer_2.Mode := #Cnv_Buffer_3.Mode := 3;// Auto Mode
           #VTD.Instruction.Enable :=
           #Extrator_Conveyor.Enabled :=
           #Cnv_Buffer_11.Instruction.Enable :=
           #Cnv_Buffer_21.Instruction.Enable :=
           #Cnv_Buffer_31.Instruction.Enable :=
           #Cnv_Buffer_41.Instruction.Enable :=
           #Cnv_Buffer_51.Instruction.Enable :=
           #Cnv_Buffer_61.Instruction.Enable :=
           #Cnv_Buffer_71.Instruction.Enable :=
           #Cnv_Buffer_81.Instruction.Enable :=
           #Cnv_Buffer_12.Instruction.Enable :=
           #Cnv_Buffer_22.Instruction.Enable :=
           #Cnv_Buffer_32.Instruction.Enable :=
           #Cnv_Buffer_42.Instruction.Enable :=
           #Cnv_Buffer_52.Instruction.Enable :=
           #Cnv_Buffer_62.Instruction.Enable :=
           #Cnv_Buffer_72.Instruction.Enable :=
           #Cnv_Buffer_82.Instruction.Enable := TRUE;
       END_IF;
       //Disable Devices in Auto/Man Mode
          #F_AutoMode(CLK:=#System.Auto_Man);

          IF #F_AutoMode.Q THEN
              #VTD.Instruction.Enable :=
              #Extrator_Conveyor.Enabled :=
              #Cnv_Buffer_11.Instruction.Enable :=
              #Cnv_Buffer_21.Instruction.Enable :=
              #Cnv_Buffer_31.Instruction.Enable :=
              #Cnv_Buffer_41.Instruction.Enable :=
              #Cnv_Buffer_51.Instruction.Enable :=
              #Cnv_Buffer_61.Instruction.Enable :=
              #Cnv_Buffer_71.Instruction.Enable :=
              #Cnv_Buffer_81.Instruction.Enable :=
              #Cnv_Buffer_12.Instruction.Enable :=
              #Cnv_Buffer_22.Instruction.Enable :=
              #Cnv_Buffer_32.Instruction.Enable :=
              #Cnv_Buffer_42.Instruction.Enable :=
              #Cnv_Buffer_52.Instruction.Enable :=
              #Cnv_Buffer_62.Instruction.Enable :=
              #Cnv_Buffer_72.Instruction.Enable :=
              #Cnv_Buffer_82.Instruction.Enable := FALSE;
          END_IF;
   END_REGION

   REGION VTD
       //VTD 
       IF #System.OrderTable[1].StepNo <> 0
           AND #System.OrderTable[1].Device = #VTD_DEVICE
           AND #System.OrderTable[1].Status = #QUEUED_STATUS
           AND NOT (#OPC_UA_State_VTD > 0 AND #OPC_UA_State_VTD < 400)
           AND NOT (#OPC_UA_State_CNV > 0 AND #OPC_UA_State_CNV < 400)
           AND NOT (#OPC_UA_State_Shuttle > 0 AND #OPC_UA_State_Shuttle < 400)
           AND NOT #System.Error
           AND NOT #Canceling
       THEN
           #VTD_CurrentOrder := 1;
       END_IF;
       IF #System.OrderTable[#VTD_CurrentOrder].StepNo <> 0
           AND #System.OrderTable[#VTD_CurrentOrder].Device = #VTD_DEVICE
           AND #System.OrderTable[#VTD_CurrentOrder].Status = #QUEUED_STATUS
           AND NOT (#OPC_UA_State_VTD > 0 AND #OPC_UA_State_VTD < 400)
           AND NOT (#OPC_UA_State_CNV > 0 AND #OPC_UA_State_CNV < 400)
           AND NOT (#OPC_UA_State_Shuttle > 0 AND #OPC_UA_State_Shuttle < 400)
           AND NOT #System.Error
           AND NOT #Canceling
       THEN

           //OPC Commands to Move VTD between floors
           // WCS => Order Table => OPC Ua Control Table

           "Control_DB".WCS_OPC_Control[#System.Id].Task_Data_Available:= TRUE; // Send the Task Data Available from WCS 
           "Control_DB".WCS_OPC_Control[#System.Id].Task_Type:= #System.OrderTable[#VTD_CurrentOrder].OPC_Control.Task_Type; // Send the Task Type - VTD = Task Type = 1
           "Control_DB".WCS_OPC_Control[#System.Id].Pallet_Type:= #System.OrderTable[#VTD_CurrentOrder].OPC_Control.Pallet_Type; // Send the Pallet Type -C=Chep/E=Euro
           "Control_DB".WCS_OPC_Control[#System.Id].Task_ID:=#System.OrderTable[#VTD_CurrentOrder].OPC_Control.Task_ID; // Send the Task ID number;
           "Control_DB".WCS_OPC_Control[#System.Id].Task_Metadata:=#System.OrderTable[#VTD_CurrentOrder].OPC_Control.Task_Metadata; // Send the Task Metadata Unique identifier
           "Control_DB".WCS_OPC_Control[#System.Id].Destination_Location:= #System.OrderTable[#VTD_CurrentOrder].OPC_Control.Destination_Location; // Send the VTD Destination Location
           "Control_DB".WCS_OPC_Control[#System.Id].Source_Location := 0; // Send the VTD Destination Location
           "Control_DB".WCS_OPC_Control[#System.Id].Pallet_Weight := #System.OrderTable[#VTD_CurrentOrder].OPC_Control.Pallet_Weight;
           #VTD_WatchdogStart := TRUE;
       END_IF;

       //RUNNING
       IF #VTD.Running AND #System.Auto_Man THEN
           #System.OrderTable[#VTD_CurrentOrder].Status := #RUNNING_STATUS;
           // "Control_DB"."Order Table"[#System.Id].Task_Data_Available := FALSE; // Send the Task Data Available from WCS 
       END_IF;

       //Cancel order
       IF #Canceling AND NOT #VTD.Running AND #VTD_CurrentOrder <> 0 THEN
           #System.OrderTable[#VTD_CurrentOrder].Status := #CANCELED_STATUS;
           #System.OrderTable[#VTD_CurrentOrder].CompleteTime := #CurrentTime;
           #VTD_CurrentOrder := 0;
           "Control_DB".WCS_OPC_Control[#System.Id].Task_Data_Available := FALSE; // Send the Task Data Available from WCS 
           "Control_DB".WCS_OPC_Control[#System.Id].Task_Type := 0; // Send the Task Type - VTD = Task Type = 1
           "Control_DB".WCS_OPC_Control[#System.Id].Pallet_Type := ' '; // Send the Pallet Type -C=Chep/E=Euro
           "Control_DB".WCS_OPC_Control[#System.Id].Task_ID := 0; // Send the Task ID number;
           "Control_DB".WCS_OPC_Control[#System.Id].Task_Metadata := ''; // Send the Task Metadata Unique identifier
           "Control_DB".WCS_OPC_Control[#System.Id].Destination_Location := 0; // Send the VTD Destination Location
           "Control_DB".WCS_OPC_Control[#System.Id].Source_Location := 0; // Send the VTD Destination 
           "Control_DB".WCS_OPC_Control[#System.Id].Pallet_Weight := 0;
       END_IF;

       //Error
       IF #VTD.Error THEN
           "Control_DB".WCS_OPC_Control[#System.Id].Task_Data_Available := FALSE; // Send the Task Data Available from WCS 
           "Control_DB".WCS_OPC_Control[#System.Id].Task_Type := 0; // Send the Task Type - VTD = Task Type = 1
           "Control_DB".WCS_OPC_Control[#System.Id].Pallet_Type := ' '; // Send the Pallet Type -C=Chep/E=Euro
           "Control_DB".WCS_OPC_Control[#System.Id].Task_ID := 0; // Send the Task ID number;
           "Control_DB".WCS_OPC_Control[#System.Id].Task_Metadata := ''; // Send the Task Metadata Unique identifier
           "Control_DB".WCS_OPC_Control[#System.Id].Destination_Location := 0; // Send the VTD Destination Location
           "Control_DB".WCS_OPC_Control[#System.Id].Source_Location := 0; // Send the VTD Destination 
           "Control_DB".WCS_OPC_Control[#System.Id].Pallet_Weight := 0;
           #System.OrderTable[#VTD_CurrentOrder].ErrorID := #VTD.VTD_Errors.Error_Word_1;
       END_IF;

       //MOVEMENT FINALIZED
       #VTDDoneRTrig(CLK := "Control_DB".WCS_OPC_Control[#System.Id].Movement_Request_Complete );
       IF #VTDDoneRTrig.Q THEN
           #VTD_WatchdogStart := FALSE;
           #System.OrderTable[#VTD_CurrentOrder].Status := #COMPLETED_STATUS;
           #System.OrderTable[#VTD_CurrentOrder].CompleteTime := #CurrentTime;
           #VTD_CurrentOrder := 0;
       END_IF;
   END_REGION
   ///////////////////////////////////////////////////////////////////////////////////////////////////////////////////////////////////////
   ///////////////////////////////////////////////////////////////////////////////////////////////////////////////////////////////////////
   REGION Pallet_InOut - Conveyors
       //VTD 
       IF #System.OrderTable[1].StepNo <> 0
           AND #System.OrderTable[1].Device = #PALLET_INOUT_DEVICE
           AND #System.OrderTable[1].Status = #QUEUED_STATUS
           AND NOT (#OPC_UA_State_CNV > 0 AND #OPC_UA_State_CNV < 400)
           AND NOT (#OPC_UA_State_VTD > 0 AND #OPC_UA_State_VTD < 400)
           AND NOT (#OPC_UA_State_Shuttle > 0 AND #OPC_UA_State_Shuttle < 400)
           AND NOT #System.Error
           AND NOT #Canceling
       THEN
           #Pallet_InOut_CurrentOrder := 1;
       END_IF;
       IF #System.OrderTable[#Pallet_InOut_CurrentOrder].StepNo <> 0
           AND #System.OrderTable[#Pallet_InOut_CurrentOrder].Device = #PALLET_INOUT_DEVICE
           AND #System.OrderTable[#Pallet_InOut_CurrentOrder].Status = #QUEUED_STATUS
           AND NOT (#OPC_UA_State_CNV > 0 AND #OPC_UA_State_CNV < 400)
           AND NOT (#OPC_UA_State_VTD > 0 AND #OPC_UA_State_VTD < 400)
           AND NOT (#OPC_UA_State_Shuttle > 0 AND #OPC_UA_State_Shuttle < 400)
           AND NOT #System.Error
           AND NOT #Canceling
       THEN
           //OPC Commands to Move Pallets IN/OUT (Buffer conveyors/Extractor conveyors)
           // WCS => Order Table => OPC Ua Control Table
           "Control_DB".WCS_OPC_Control[#System.Id].Task_Data_Available := TRUE; // Send the Task Data Available from WCS 
           "Control_DB".WCS_OPC_Control[#System.Id].Task_Type := #System.OrderTable[#Pallet_InOut_CurrentOrder].OPC_Control.Task_Type; // Send the Task Type - Pallet Transfer IN/OUT = Task Type = 4/
           "Control_DB".WCS_OPC_Control[#System.Id].Task_ID := #System.OrderTable[#Pallet_InOut_CurrentOrder].OPC_Control.Task_ID; // Send the Task ID number;
           "Control_DB".WCS_OPC_Control[#System.Id].Task_Metadata := #System.OrderTable[#Pallet_InOut_CurrentOrder].OPC_Control.Task_Metadata; // Send the Task Metadata Unique identifier
           "Control_DB".WCS_OPC_Control[#System.Id].Source_Location := #System.OrderTable[#Pallet_InOut_CurrentOrder].OPC_Control.Source_Location; // Send the Source Location from the Conveyor
           "Control_DB".WCS_OPC_Control[#System.Id].Destination_Location := #System.OrderTable[#Pallet_InOut_CurrentOrder].OPC_Control.Destination_Location; // Send the Destination Location to the Conveyor;
           "Control_DB".WCS_OPC_Control[#System.Id].Pallet_Type := #System.OrderTable[#Pallet_InOut_CurrentOrder].OPC_Control.Pallet_Type;
           "Control_DB".WCS_OPC_Control[#System.Id].Pallet_Alignment := #System.OrderTable[#Pallet_InOut_CurrentOrder].OPC_Control.Pallet_Alignment;
           #Pallet_InOut_WatchdogStart := TRUE;
       END_IF;

       //RUNNING
       // IF (#Extrator_Conveyor.Running OR #Cnv_Buffer_11.Running OR #Cnv_Buffer_21.Running OR #Cnv_Buffer_31.Running OR #Cnv_Buffer_41.Running OR #Cnv_Buffer_51.Running OR #Cnv_Buffer_61.Running OR #Cnv_Buffer_71.Running OR #Cnv_Buffer_81.Running
       //     OR #Cnv_Buffer_12.Running OR #Cnv_Buffer_22.Running OR #Cnv_Buffer_32.Running OR #Cnv_Buffer_42.Running OR #Cnv_Buffer_52.Running OR #Cnv_Buffer_62.Running OR #Cnv_Buffer_72.Running OR #Cnv_Buffer_82.Running)
       //     AND #System.Auto_Man THEN
       IF #OPC_UA_State_CNV > 0 AND #OPC_UA_State_CNV < 400
           AND #System.Auto_Man THEN
           #System.OrderTable[#Pallet_InOut_CurrentOrder].Status := #RUNNING_STATUS;
       END_IF;

       //Cancel order
       IF #Canceling AND NOT (#Extrator_Conveyor.Running OR #Cnv_Buffer_11.Running OR #Cnv_Buffer_21.Running OR #Cnv_Buffer_31.Running OR #Cnv_Buffer_41.Running OR #Cnv_Buffer_51.Running OR #Cnv_Buffer_61.Running OR #Cnv_Buffer_71.Running OR #Cnv_Buffer_81.Running
           OR #Cnv_Buffer_12.Running OR #Cnv_Buffer_22.Running OR #Cnv_Buffer_32.Running OR #Cnv_Buffer_42.Running OR #Cnv_Buffer_52.Running OR #Cnv_Buffer_62.Running OR #Cnv_Buffer_72.Running OR #Cnv_Buffer_82.Running)
           AND #Pallet_InOut_CurrentOrder <> 0 THEN
           #System.OrderTable[#Pallet_InOut_CurrentOrder].Status := #CANCELED_STATUS;
           #System.OrderTable[#Pallet_InOut_CurrentOrder].CompleteTime := #CurrentTime;
           #Pallet_InOut_CurrentOrder := 0;
           "Control_DB".WCS_OPC_Control[#System.Id].Task_Data_Available := FALSE; // Send the Task Data Available from WCS 
           "Control_DB".WCS_OPC_Control[#System.Id].Task_Type := #System.OrderTable[#Pallet_InOut_CurrentOrder].OPC_Control.Task_Type; // Send the Task Type - Pallet Transfer IN/OUT = Task Type = 4/
           "Control_DB".WCS_OPC_Control[#System.Id].Task_ID := #System.OrderTable[#Pallet_InOut_CurrentOrder].OPC_Control.Task_ID; // Send the Task ID number;
           "Control_DB".WCS_OPC_Control[#System.Id].Task_Metadata := #System.OrderTable[#Pallet_InOut_CurrentOrder].OPC_Control.Task_Metadata; // Send the Task Metadata Unique identifier
           "Control_DB".WCS_OPC_Control[#System.Id].Source_Location := #System.OrderTable[#Pallet_InOut_CurrentOrder].OPC_Control.Source_Location; // Send the Source Location from the Conveyor
           "Control_DB".WCS_OPC_Control[#System.Id].Destination_Location := #System.OrderTable[#Pallet_InOut_CurrentOrder].OPC_Control.Destination_Location; // Send the Destination Location to the Conveyor;
           "Control_DB".WCS_OPC_Control[#System.Id].Pallet_Type := #System.OrderTable[#Pallet_InOut_CurrentOrder].OPC_Control.Pallet_Type;
           "Control_DB".WCS_OPC_Control[#System.Id].Pallet_Alignment := #System.OrderTable[#Pallet_InOut_CurrentOrder].OPC_Control.Pallet_Alignment;
       END_IF;

       //Error
       IF (#Extrator_Conveyor.Error OR #Cnv_Buffer_11.Error OR #Cnv_Buffer_21.Error OR #Cnv_Buffer_31.Error OR #Cnv_Buffer_41.Error OR #Cnv_Buffer_51.Error OR #Cnv_Buffer_61.Error OR #Cnv_Buffer_71.Error OR #Cnv_Buffer_81.Error
           OR #Cnv_Buffer_12.Error OR #Cnv_Buffer_22.Error OR #Cnv_Buffer_32.Error OR #Cnv_Buffer_42.Error OR #Cnv_Buffer_52.Error OR #Cnv_Buffer_62.Error OR #Cnv_Buffer_72.Error OR #Cnv_Buffer_82.Error) THEN
           "Control_DB".WCS_OPC_Control[#System.Id].Task_Data_Available := FALSE; // Send the Task Data Available from WCS 
           "Control_DB".WCS_OPC_Control[#System.Id].Task_Type := #System.OrderTable[#Pallet_InOut_CurrentOrder].OPC_Control.Task_Type; // Send the Task Type - Pallet Transfer IN/OUT = Task Type = 4/
           "Control_DB".WCS_OPC_Control[#System.Id].Task_ID := #System.OrderTable[#Pallet_InOut_CurrentOrder].OPC_Control.Task_ID; // Send the Task ID number;
           "Control_DB".WCS_OPC_Control[#System.Id].Task_Metadata := #System.OrderTable[#Pallet_InOut_CurrentOrder].OPC_Control.Task_Metadata; // Send the Task Metadata Unique identifier
           "Control_DB".WCS_OPC_Control[#System.Id].Source_Location := #System.OrderTable[#Pallet_InOut_CurrentOrder].OPC_Control.Source_Location; // Send the Source Location from the Conveyor
           "Control_DB".WCS_OPC_Control[#System.Id].Destination_Location := #System.OrderTable[#Pallet_InOut_CurrentOrder].OPC_Control.Destination_Location; // Send the Destination Location to the Conveyor;
           "Control_DB".WCS_OPC_Control[#System.Id].Pallet_Type := #System.OrderTable[#Pallet_InOut_CurrentOrder].OPC_Control.Pallet_Type;
           "Control_DB".WCS_OPC_Control[#System.Id].Pallet_Alignment := #System.OrderTable[#Pallet_InOut_CurrentOrder].OPC_Control.Pallet_Alignment;
           #System.OrderTable[#Pallet_InOut_CurrentOrder].Status := #ERROR_STATUS;

           // #System.OrderTable[#Pallet_InOut_CurrentOrder].ErrorID := (#Extrator_Conveyor.Cnv_Errors. OR #Cnv_Buffer_11.Error OR #Cnv_Buffer_21.Error OR #Cnv_Buffer_31.Error OR #Cnv_Buffer_41.Error OR #Cnv_Buffer_51.Error OR #Cnv_Buffer_61.Error OR #Cnv_Buffer_71.Error OR #Cnv_Buffer_81.Error
           // OR #Cnv_Buffer_12.Error OR #Cnv_Buffer_22.Error OR #Cnv_Buffer_32.Error OR #Cnv_Buffer_42.Error OR #Cnv_Buffer_52.Error OR #Cnv_Buffer_62.Error OR #Cnv_Buffer_72.Error OR #Cnv_Buffer_82.Error);
       END_IF;

       //MOVEMENT FINALIZED
       #Pallet_InOut_RTrig(CLK := "Control_DB".WCS_OPC_Control[#System.Id].Movement_Request_Complete);
       IF #Pallet_InOut_RTrig.Q THEN
           "Control_DB".WCS_OPC_Control[#System.Id].Task_Data_Available := FALSE; //#System.OrderTable[#Pallet_InOut_CurrentOrder].OPC_Control.Task_Data_Available; // Send the Task Data Available from WCS 
           "Control_DB".WCS_OPC_Control[#System.Id].Task_Type := #System.OrderTable[#Pallet_InOut_CurrentOrder].OPC_Control.Task_Type; // Send the Task Type - Pallet Transfer IN/OUT = Task Type = 4/
           "Control_DB".WCS_OPC_Control[#System.Id].Task_ID := #System.OrderTable[#Pallet_InOut_CurrentOrder].OPC_Control.Task_ID; // Send the Task ID number;
           "Control_DB".WCS_OPC_Control[#System.Id].Task_Metadata := #System.OrderTable[#Pallet_InOut_CurrentOrder].OPC_Control.Task_Metadata; // Send the Task Metadata Unique identifier
           "Control_DB".WCS_OPC_Control[#System.Id].Source_Location := #System.OrderTable[#Pallet_InOut_CurrentOrder].OPC_Control.Source_Location; // Send the Source Location from the Conveyor
           "Control_DB".WCS_OPC_Control[#System.Id].Destination_Location := #System.OrderTable[#Pallet_InOut_CurrentOrder].OPC_Control.Destination_Location; // Send the Destination Location to the Conveyor;
           "Control_DB".WCS_OPC_Control[#System.Id].Pallet_Type := #System.OrderTable[#Pallet_InOut_CurrentOrder].OPC_Control.Pallet_Type;
           "Control_DB".WCS_OPC_Control[#System.Id].Pallet_Alignment := #System.OrderTable[#Pallet_InOut_CurrentOrder].OPC_Control.Pallet_Alignment;
           #System.OrderTable[#Pallet_InOut_CurrentOrder].Status := #COMPLETED_STATUS;
           #System.OrderTable[#Pallet_InOut_CurrentOrder].CompleteTime := #CurrentTime;
           #Pallet_InOut_CurrentOrder := 0;
       END_IF;
   END_REGION
   ///////////////////////////////////////////////////////////////////////////////////////////////////////////////////////////////////////
   ///////////////////////////////////////////////////////////////////////////////////////////////////////////////////////////////////////
   REGION Shuttle_InOut
       //Shuttle Interlock on VTD 
       IF #System.OrderTable[1].StepNo <> 0
           AND #System.OrderTable[1].Device = #SHUTTLE_INOUT_DEVICE
           AND #System.OrderTable[1].Status = #QUEUED_STATUS
           AND NOT (#OPC_UA_State_Shuttle > 0 AND #OPC_UA_State_Shuttle < 400)
           AND NOT (#OPC_UA_State_CNV > 0 AND #OPC_UA_State_CNV < 400)
           AND NOT (#OPC_UA_State_VTD > 0 AND #OPC_UA_State_VTD < 400)
           AND NOT #System.Error
           AND NOT #Canceling
       THEN
           #Shuttle_InOut_CurrentOrder := 1;
       END_IF;
       IF #System.OrderTable[#Shuttle_InOut_CurrentOrder].StepNo <> 0
           AND #System.OrderTable[#Shuttle_InOut_CurrentOrder].Device = #SHUTTLE_INOUT_DEVICE
           AND #System.OrderTable[#Shuttle_InOut_CurrentOrder].Status = #QUEUED_STATUS
           AND NOT (#OPC_UA_State_Shuttle > 0 AND #OPC_UA_State_Shuttle < 400)
           AND NOT (#OPC_UA_State_CNV > 0 AND #OPC_UA_State_CNV < 400)
           AND NOT (#OPC_UA_State_VTD > 0 AND #OPC_UA_State_VTD < 400)
           AND NOT #System.Error
           AND NOT #Canceling
       THEN
           //OPC Commands to Move Shuttle IN/OUT (Shuttles IN/OUT)
           // WCS => Order Table => OPC Ua Control Table
           "Control_DB".WCS_OPC_Control[#System.Id].Task_Data_Available := TRUE;// Send the Task Data Available from WCS
           "Control_DB".WCS_OPC_Control[#System.Id].Task_ID := #System.OrderTable[#Shuttle_InOut_CurrentOrder].OPC_Control.Task_ID; // Send the Task ID number;
           "Control_DB".WCS_OPC_Control[#System.Id].Task_Metadata := #System.OrderTable[#Shuttle_InOut_CurrentOrder].OPC_Control.Task_Metadata; // Send the Task Metadata Unique identifier
           "Control_DB".WCS_OPC_Control[#System.Id].Pallet_Type := #System.OrderTable[#Shuttle_InOut_CurrentOrder].OPC_Control.Pallet_Type; // Send Pallet Type
           "Control_DB".WCS_OPC_Control[#System.Id].Task_Type := #System.OrderTable[#Shuttle_InOut_CurrentOrder].OPC_Control.Task_Type; // Send the Task Type - Pallet Transfer IN/OUT = Task Type = 4/
           "Control_DB".WCS_OPC_Control[#System.Id].Shuttle_ID := #System.OrderTable[#Shuttle_InOut_CurrentOrder].OPC_Control.Shuttle_ID;// Send the Shuttle ID
           "Control_DB".WCS_OPC_Control[#System.Id].Shuttle_Loaded := #System.OrderTable[#Shuttle_InOut_CurrentOrder].OPC_Control.Shuttle_Loaded; // Send the Shuttle status (Loaded/Unloaded)
           "Control_DB".WCS_OPC_Control[#System.Id].Source_Location := #System.OrderTable[#Shuttle_InOut_CurrentOrder].OPC_Control.Source_Location; // Send the Source Location from the Conveyor
           "Control_DB".WCS_OPC_Control[#System.Id].Destination_Location := #System.OrderTable[#Shuttle_InOut_CurrentOrder].OPC_Control.Destination_Location; // Send the Destination Location to the Conveyor;
           #Shuttle_InOut_WatchdogStart := TRUE;
       END_IF;

       //RUNNING
       IF #OPC_UA_State_Shuttle > 0 AND #OPC_UA_State_Shuttle < 400 AND #System.Auto_Man THEN
           #System.OrderTable[#Shuttle_InOut_CurrentOrder].Status := #RUNNING_STATUS;
       END_IF;

       //Cancel order
       IF #Canceling AND NOT (#VTD.Running) AND #Shuttle_InOut_CurrentOrder <> 0 THEN
           #System.OrderTable[#Shuttle_InOut_CurrentOrder].Status := #CANCELED_STATUS;
           #System.OrderTable[#Shuttle_InOut_CurrentOrder].CompleteTime := #CurrentTime;
           #Shuttle_InOut_CurrentOrder := 0;
           "Control_DB".WCS_OPC_Control[#System.Id].Task_Data_Available := FALSE;// Send the Task Data Available from WCS 
           "Control_DB".WCS_OPC_Control[#System.Id].Task_ID := #System.OrderTable[#Shuttle_InOut_CurrentOrder].OPC_Control.Task_ID; // Send the Task ID number;
           "Control_DB".WCS_OPC_Control[#System.Id].Task_Metadata := #System.OrderTable[#Shuttle_InOut_CurrentOrder].OPC_Control.Task_Metadata; // Send the Task Metadata Unique identifier
           "Control_DB".WCS_OPC_Control[#System.Id].Pallet_Type := #System.OrderTable[#Shuttle_InOut_CurrentOrder].OPC_Control.Pallet_Type; // Send Pallet Type
           "Control_DB".WCS_OPC_Control[#System.Id].Task_Type := #System.OrderTable[#Shuttle_InOut_CurrentOrder].OPC_Control.Task_Type; // Send the Task Type - Pallet Transfer IN/OUT = Task Type = 4/
           "Control_DB".WCS_OPC_Control[#System.Id].Shuttle_ID := #System.OrderTable[#Shuttle_InOut_CurrentOrder].OPC_Control.Shuttle_ID;// Send the Shuttle ID
           "Control_DB".WCS_OPC_Control[#System.Id].Shuttle_Loaded := #System.OrderTable[#Shuttle_InOut_CurrentOrder].OPC_Control.Shuttle_Loaded; // Send the Shuttle status (Loaded/Unloaded)
           "Control_DB".WCS_OPC_Control[#System.Id].Source_Location := #System.OrderTable[#Shuttle_InOut_CurrentOrder].OPC_Control.Source_Location; // Send the Source Location from the Conveyor
           "Control_DB".WCS_OPC_Control[#System.Id].Destination_Location := #System.OrderTable[#Shuttle_InOut_CurrentOrder].OPC_Control.Destination_Location; // Send the Destination Location to the Conveyor;
       END_IF;

       //Error
       IF #OPC_UA_State_Shuttle = 400 THEN
           "Control_DB".WCS_OPC_Control[#System.Id].Task_Data_Available := FALSE;//#System.OrderTable[#Shuttle_InOut_CurrentOrder].OPC_Control.Task_Data_Available; // Send the Task Data Available from WCS 
           "Control_DB".WCS_OPC_Control[#System.Id].Task_ID := #System.OrderTable[#Shuttle_InOut_CurrentOrder].OPC_Control.Task_ID; // Send the Task ID number;
           "Control_DB".WCS_OPC_Control[#System.Id].Task_Metadata := #System.OrderTable[#Shuttle_InOut_CurrentOrder].OPC_Control.Task_Metadata; // Send the Task Metadata Unique identifier
           "Control_DB".WCS_OPC_Control[#System.Id].Pallet_Type := #System.OrderTable[#Shuttle_InOut_CurrentOrder].OPC_Control.Pallet_Type; // Send Pallet Type
           "Control_DB".WCS_OPC_Control[#System.Id].Task_Type := #System.OrderTable[#Shuttle_InOut_CurrentOrder].OPC_Control.Task_Type; // Send the Task Type - Pallet Transfer IN/OUT = Task Type = 4/
           "Control_DB".WCS_OPC_Control[#System.Id].Shuttle_ID := #System.OrderTable[#Shuttle_InOut_CurrentOrder].OPC_Control.Shuttle_ID;// Send the Shuttle ID
           "Control_DB".WCS_OPC_Control[#System.Id].Shuttle_Loaded := #System.OrderTable[#Shuttle_InOut_CurrentOrder].OPC_Control.Shuttle_Loaded; // Send the Shuttle status (Loaded/Unloaded)
           "Control_DB".WCS_OPC_Control[#System.Id].Source_Location := #System.OrderTable[#Shuttle_InOut_CurrentOrder].OPC_Control.Source_Location; // Send the Source Location from the Conveyor
           "Control_DB".WCS_OPC_Control[#System.Id].Destination_Location := #System.OrderTable[#Shuttle_InOut_CurrentOrder].OPC_Control.Destination_Location; // Send the Destination Location to the Conveyor;
           #System.OrderTable[#Shuttle_InOut_CurrentOrder].Status := #ERROR_STATUS;
           #System.OrderTable[#Shuttle_InOut_CurrentOrder].ErrorID := (#VTD.VTD_Errors.Error_Word_3);
       END_IF;

       //MOVEMENT FINALIZED
       #Shuttle_InOut_RTrig(CLK := #VTD.Shuttle_Interlock.Interlock_Complete);
       IF #Shuttle_InOut_RTrig.Q THEN
           "Control_DB".WCS_OPC_Control[#System.Id].Task_Data_Available := FALSE;//#System.OrderTable[#Shuttle_InOut_CurrentOrder].OPC_Control.Task_Data_Available; // Send the Task Data Available from WCS 
           "Control_DB".WCS_OPC_Control[#System.Id].Task_ID := #System.OrderTable[#Shuttle_InOut_CurrentOrder].OPC_Control.Task_ID; // Send the Task ID number;
           "Control_DB".WCS_OPC_Control[#System.Id].Task_Metadata := #System.OrderTable[#Shuttle_InOut_CurrentOrder].OPC_Control.Task_Metadata; // Send the Task Metadata Unique identifier
           "Control_DB".WCS_OPC_Control[#System.Id].Pallet_Type := #System.OrderTable[#Shuttle_InOut_CurrentOrder].OPC_Control.Pallet_Type; // Send Pallet Type
           "Control_DB".WCS_OPC_Control[#System.Id].Task_Type := #System.OrderTable[#Shuttle_InOut_CurrentOrder].OPC_Control.Task_Type; // Send the Task Type - Pallet Transfer IN/OUT = Task Type = 4/
           "Control_DB".WCS_OPC_Control[#System.Id].Shuttle_ID := #System.OrderTable[#Shuttle_InOut_CurrentOrder].OPC_Control.Shuttle_ID;// Send the Shuttle ID
           "Control_DB".WCS_OPC_Control[#System.Id].Shuttle_Loaded := #System.OrderTable[#Shuttle_InOut_CurrentOrder].OPC_Control.Shuttle_Loaded; // Send the Shuttle status (Loaded/Unloaded)
           "Control_DB".WCS_OPC_Control[#System.Id].Source_Location := #System.OrderTable[#Shuttle_InOut_CurrentOrder].OPC_Control.Source_Location; // Send the Source Location from the Conveyor
           "Control_DB".WCS_OPC_Control[#System.Id].Destination_Location := #System.OrderTable[#Shuttle_InOut_CurrentOrder].OPC_Control.Destination_Location; // Send the Destination Location to the Conveyor;

           #Shuttle_InOut_WatchdogStart := FALSE;
           #System.OrderTable[#Shuttle_InOut_CurrentOrder].Status := #COMPLETED_STATUS;
           #System.OrderTable[#Shuttle_InOut_CurrentOrder].CompleteTime := #CurrentTime;
           #Shuttle_InOut_CurrentOrder := 0;
       END_IF;
   END_REGION
   ///////////////////////////////////////////////////////////////////////////////////////////////////////////////////////////////////////
   ///////////////////////////////////////////////////////////////////////////////////////////////////////////////////////////////////////

   REGION Max Running Order Number
       #MaxRunningOrderNo := MAX(IN1 := #VTD_CurrentOrder, IN2 := #Pallet_InOut_CurrentOrder,
                                 IN3 := #Shuttle_InOut_CurrentOrder, IN4 := #System.CurrentOrder);

   END_REGION

   REGION Pause Orders
       #ErrorRTrig(CLK := #System.Error);
       #PauseRTrig(CLK := #System.PauseOrders OR NOT #System.Auto_Man);
       IF #ErrorRTrig.Q OR #PauseRTrig.Q THEN
           #System.PauseOrders := FALSE;
           #System.Paused := #MaxRunningOrderNo > 0;
           IF #System.Paused THEN
               FOR #i := 1 TO UDINT_TO_DINT(#MaxRunningOrderNo) DO
                   IF #System.OrderTable[#i].Status = '' THEN
                       EXIT;
                   ELSIF #System.OrderTable[#i].Status = #QUEUED_STATUS THEN
                       #System.OrderTable[#i].Status := #PAUSED_STATUS;
                   ELSIF #System.OrderTable[#i].Status = #RUNNING_STATUS AND NOT #System.Auto_Man THEN
                       #System.OrderTable[#i].Status := #CANCELED_STATUS;
                   END_IF;
               END_FOR;
           END_IF;
       END_IF;
       IF #System.Paused AND #MaxRunningOrderNo = 0 THEN
           #System.Paused := FALSE;
       END_IF;
   END_REGION

   REGION Cancel Orders
       #CancelRTrig(CLK := #System.CancelOrders);
       (*#WeighingStation.Cancel := #ProfileStation.Cancel:= #CancelRTrig.Q*);
       IF #CancelRTrig.Q THEN
           #Canceling := TRUE;
           #System.CancelOrders := FALSE;
           #System.Paused := FALSE;
           FOR #i := 1 TO UDINT_TO_DINT(#MaxRunningOrderNo) DO
               IF #System.OrderTable[#i].Status = '' THEN
                   CONTINUE;
               ELSIF #System.OrderTable[#i].Status = #PAUSED_STATUS
                   OR #System.OrderTable[#i].Status = #QUEUED_STATUS
               THEN
                   #System.OrderTable[#i].Status := #CANCELED_STATUS;
                   #System.OrderTable[#i].CompleteTime := #CurrentTime;
               ELSIF #System.OrderTable[#i].Status = #ERROR_STATUS
               THEN
                   #System.OrderTable[#i].Status := #ERROR_CANCELED_STATUS;
                   #System.OrderTable[#i].CompleteTime := #CurrentTime;
               END_IF;
           END_FOR;
           #System.CurrentOrder := 0;
       END_IF;
       IF #Canceling AND NOT (#VTD.Running OR #Extrator_Conveyor.Running OR #Cnv_Buffer_11.Running OR #Cnv_Buffer_21.Running OR #Cnv_Buffer_41.Running) THEN
           #Canceling := FALSE;
           #VTD_CurrentOrder := #Pallet_InOut_CurrentOrder:= #Shuttle_InOut_CurrentOrder := 0;
       END_IF;
   END_REGION

   REGION Resume Orders
       #ResumeRTrig(CLK := #System.ResumeOrders);
       IF #ResumeRTrig.Q THEN
           #System.ResumeOrders := FALSE;
           #System.CurrentOrder := #MaxRunningOrderNo;
           IF NOT #System.Error THEN
               #System.Paused := FALSE;
               FOR #i := 1 TO UDINT_TO_DINT(#MaxRunningOrderNo) DO
                   IF #System.OrderTable[#i].Status = '' THEN
                       EXIT;
                   ELSIF #System.OrderTable[#i].Status = #PAUSED_STATUS
                       OR #System.OrderTable[#i].Status = #ERROR_STATUS
                   THEN
                       #System.OrderTable[#i].Status := #QUEUED_STATUS;
                   END_IF;
               END_FOR;
           END_IF;

       END_IF;
   END_REGION

   REGION Order Handler
       IF #System.Running AND NOT #System.Error
           AND (#System.OrderTable[#System.CurrentOrder].Status = #COMPLETED_STATUS
           OR #System.OrderTable[#System.CurrentOrder].Status = #ERROR_STATUS
           OR #System.OrderTable[#System.CurrentOrder].Status = #ERROR_CANCELED_STATUS
           OR #System.OrderTable[#System.CurrentOrder].Sequence = 0)
       THEN
           IF #System.CurrentOrder > 0 THEN
               #System.CurrentOrder -= 1;
           ELSE
               #System.CurrentOrder := 0;
           END_IF;
       END_IF;
   END_REGION

   REGION Watchdogs
       //Watchdog Timers

       #VTD_WatchdogTimer(IN := #VTD_WatchdogStart,
                          PT := UDINT_TO_TIME(#Watchdog.VTD * 60000),
                          Q => #System.Watchdog_TimeOut.VTD);
       #Pallet_InOut_WatchdogTimer(IN := #Pallet_InOut_WatchdogStart,
                                   PT := UDINT_TO_TIME(#Watchdog.Pallet_INOut * 60000),
                                   Q => #System.Watchdog_TimeOut.Pallet_InOut);
       #Shuttle_InOut_WatchdogTimer(IN := #Shuttle_InOut_WatchdogStart,
                                    PT := UDINT_TO_TIME(#Watchdog.Shuttle_INOut * 60000),
                                    Q => #System.Watchdog_TimeOut.Shuttle_InOut);

   END_REGION

   REGION Reset Next Order Number
       IF #System.NextOrder > 1
           AND #CurrentDTL.HOUR = 0
           AND #CurrentDTL.MINUTE = 0
           AND #CurrentDTL.SECOND = 0
       THEN
           #System.NextOrder := 1;
       END_IF;

   END_REGION

   REGION #System Mode and State
       #System.Selected := #System_Selected; // System selected
       #System.Ready := NOT #System.Error AND #System.Selected;
       #System.Auto_Man := #AutoMan_Switch;
       #System.Running := #VTD.Running OR #Extrator_Conveyor.Running OR #Cnv_Buffer_11.Running OR #Cnv_Buffer_21.Running OR
       #Cnv_Buffer_21.Running OR #Cnv_Buffer_31.Running OR #Cnv_Buffer_41.Running OR #Cnv_Buffer_51.Running OR
       #Cnv_Buffer_61.Running OR #Cnv_Buffer_71.Running OR #Cnv_Buffer_81.Running OR #Cnv_Buffer_12.Running OR
       #Cnv_Buffer_22.Running OR #Cnv_Buffer_32.Running OR #Cnv_Buffer_42.Running OR #Cnv_Buffer_52.Running OR
       #Cnv_Buffer_62.Running OR #Cnv_Buffer_72.Running OR #Cnv_Buffer_82.Running;

       #System.Error := #VTD.Error OR #Extrator_Conveyor.Error OR #Cnv_Buffer_11.Error OR #Cnv_Buffer_21.Error OR
       #Cnv_Buffer_21.Error OR #Cnv_Buffer_31.Error OR #Cnv_Buffer_41.Error OR #Cnv_Buffer_51.Error OR
       #Cnv_Buffer_61.Error OR #Cnv_Buffer_71.Error OR #Cnv_Buffer_81.Error OR #Cnv_Buffer_12.Error OR
       #Cnv_Buffer_22.Error OR #Cnv_Buffer_32.Error OR #Cnv_Buffer_42.Error OR #Cnv_Buffer_52.Error OR
       #Cnv_Buffer_62.Error OR #Cnv_Buffer_72.Error OR #Cnv_Buffer_82.Error OR #OPC_UA_State_VTD = 400 OR #OPC_UA_State_Shuttle = 400 OR #OPC_UA_State_CNV = 400;

       #System.IDLE := NOT #System.Running AND NOT #System.Paused AND NOT #System.Error;
       IF #System.Running THEN
           #System.State := 1;
       ELSIF #System.Paused AND NOT #System.Error THEN
           #System.State := 2;
       ELSIF #System.Error THEN
           #System.State := 3;
       ELSE
           #System.State := 0;
       END_IF;
   END_REGION

   REGION Clear order table
       IF #Clear_OrderTable THEN
           FOR #i := 0 TO 99 DO
               #System.OrderTable[#i] := #EmptyOrder;
           END_FOR;
           "Control_DB".WCS_OPC_Control[#System.Id].Task_Data_Available := FALSE;
       END_IF;
   END_REGION
END_FUNCTION_BLOCK

FUNCTION "LGX_SM_FC" : Void   // FC13, SCL
{ S7_Optimized_Access := 'TRUE' }
VERSION : 0.1
// stored: AutoNumber true, IsIECCheckEnabled false, SetENOAutomatically false, UDAEnableTagReadback false
   VAR_OUTPUT
      Fault_Handshake_Infeed_1 : Bool;
      Fault_Handshake_Infeed_2 : Bool;
      Fault_Handshake_Infeed_3 : Bool;
      Fault_Handshake_Outfeed_1 : Bool;
      Fault_Handshake_Outfeed_2 : Bool;
      Fault_Handshake_Outfeed_3 : Bool;
   END_VAR
   VAR CONSTANT
      AUTO_RUNNING : UInt := 0;
   END_VAR
BEGIN
   REGION INFEED
       // 1
       "Handshake_Infeed_FC"(Infeed_Stop_Sensor := "Control_DB".LCnv_Sys[1].Cnv_Level[1].Cnv1.Inputs.Right,
                             Ready_To_Receive := "Control_DB".LCnv_Sys[1].Cnv_Level[1].Cnv1.Instruction.Inbound_Ready AND
                             NOT "Control_DB".Gate_Station[1].Requested_Access AND NOT "Control_DB".Gate_Station[2].Requested_Access,
                             Auto_Mode := "Control_DB".LCnv_Sys[1].Cnv_Level[1].Cnv1.Mode = 3,
                             Transfer_In_Progress := "Control_DB".LCnv_Sys[1].Cnv_Level[1].Cnv1.Running,
                             DB_LGX_To_SM_Infeed_Ready_To_Send := "DB_Receive_Data_From_Logistex".J1310_Conv_Infeed.LGXReadyToSend,
                             DB_LGX_To_SM_Infeed_Transfer_In_Progress := "DB_Receive_Data_From_Logistex".J1310_Conv_Infeed.LGXTransferingInProgress,
                             Fault_Handshake => #Fault_Handshake_Infeed_1,
                             DB_SM_To_LGX_Infeed_Ready_To_Receive => "DB_Send_Data_To_Logistex".VTD_J1310_INFEED.SPMReadyToReceive,
                             DB_SM_To_LGX_Infeed_Pallet_Received => "DB_Send_Data_To_Logistex".VTD_J1310_INFEED.SPMTransferingOccupied,
                             DB_SM_To_LGX_Infeed_Transfer_In_Progress => "DB_Send_Data_To_Logistex".VTD_J1310_INFEED.SPMTransferingInProgress);

       // 2
       "Handshake_Infeed_FC"(Infeed_Stop_Sensor := "Control_DB".LCnv_Sys[2].Cnv_Level[1].Cnv1.Inputs.Right,
                             Ready_To_Receive := "Control_DB".LCnv_Sys[2].Cnv_Level[1].Cnv1.Instruction.Inbound_Ready AND
                             NOT "Control_DB".Gate_Station[3].Requested_Access AND NOT "Control_DB".Gate_Station[4].Requested_Access,
                             Auto_Mode := "Control_DB".LCnv_Sys[2].Cnv_Level[1].Cnv1.Mode = 3,
                             Transfer_In_Progress := "Control_DB".LCnv_Sys[2].Cnv_Level[1].Cnv1.Running,
                             DB_LGX_To_SM_Infeed_Ready_To_Send := "DB_Receive_Data_From_Logistex".J1320_Conv_Infeed.LGXReadyToSend,
                             DB_LGX_To_SM_Infeed_Transfer_In_Progress := "DB_Receive_Data_From_Logistex".J1320_Conv_Infeed.LGXTransferingInProgress,
                             Fault_Handshake => #Fault_Handshake_Infeed_2,
                             DB_SM_To_LGX_Infeed_Ready_To_Receive => "DB_Send_Data_To_Logistex".VTD_J1320_INFEED.SPMReadyToReceive,
                             DB_SM_To_LGX_Infeed_Pallet_Received => "DB_Send_Data_To_Logistex".VTD_J1320_INFEED.SPMTransferingOccupied,
                             DB_SM_To_LGX_Infeed_Transfer_In_Progress => "DB_Send_Data_To_Logistex".VTD_J1320_INFEED.SPMTransferingInProgress);

       // 3
       "Handshake_Infeed_FC"(Infeed_Stop_Sensor := "Control_DB".LCnv_Sys[3].Cnv_Level[1].Cnv1.Inputs.Right,
                             Ready_To_Receive := "Control_DB".LCnv_Sys[3].Cnv_Level[1].Cnv1.Instruction.Inbound_Ready AND
                             NOT "Control_DB".Gate_Station[5].Requested_Access AND NOT "Control_DB".Gate_Station[6].Requested_Access,
                             Auto_Mode := "Control_DB".LCnv_Sys[3].Cnv_Level[1].Cnv1.Mode = 3,
                             Transfer_In_Progress := "Control_DB".LCnv_Sys[3].Cnv_Level[1].Cnv1.Running,
                             DB_LGX_To_SM_Infeed_Ready_To_Send := "DB_Receive_Data_From_Logistex".J1330_Conv_Infeed.LGXReadyToSend,
                             DB_LGX_To_SM_Infeed_Transfer_In_Progress := "DB_Receive_Data_From_Logistex".J1330_Conv_Infeed.LGXTransferingInProgress,
                             Fault_Handshake => #Fault_Handshake_Infeed_3,
                             DB_SM_To_LGX_Infeed_Ready_To_Receive => "DB_Send_Data_To_Logistex".VTD_J1330_INFEED.SPMReadyToReceive,
                             DB_SM_To_LGX_Infeed_Pallet_Received => "DB_Send_Data_To_Logistex".VTD_J1330_INFEED.SPMTransferingOccupied,
                             DB_SM_To_LGX_Infeed_Transfer_In_Progress => "DB_Send_Data_To_Logistex".VTD_J1330_INFEED.SPMTransferingInProgress);

   END_REGION ;

   REGION OUTFEED
       // 1
       "Handshake_Outfeed_FC"(Auto_Mode := "Control_DB".LCnv_Sys[1].Cnv_Level[1].Cnv2.Mode = 3,
                              Ready_To_Send := "Control_DB".LCnv_Sys[1].Cnv_Level[1].Cnv2.Instruction.Outbound_Ready,
                              Conv_Occupied := "Control_DB".LCnv_Sys[1].Cnv_Level[1].Cnv2.Cnv_Occupied,
                              Transfer_In_Progress := "Control_DB".LCnv_Sys[1].Cnv_Level[1].Cnv2.Running,
                              DB_LGX_To_SM_Outfeed_Ready_To_Receive := "DB_Receive_Data_From_Logistex".J1310_Conv_Oufeed.LGXReadyToReceive,
                              Fault_Handshake => #Fault_Handshake_Outfeed_1,
                              DB_SM_To_LGX_Outfeed_Transfer_In_Progress => "DB_Send_Data_To_Logistex".VTD_J1310_OUTFEED.SPMTransferingInProgress,
                              DB_SM_To_LGX_Outfeed_Ocuppied => "DB_Send_Data_To_Logistex".VTD_J1310_OUTFEED.SPMTransferingOccupied,
                              DB_SM_To_LGX_Outfeed_Ready_To_Send => "DB_Send_Data_To_Logistex".VTD_J1310_OUTFEED.SPMReadyToSend);

       // Pallet tpe
       IF "Control_DB".LCnv_Sys[1].Cnv_Level[1].Cnv2.Pallet_Type = 1 THEN
           "DB_Send_Data_To_Logistex".VTD_J1310_OUTFEED.Pallet_ID[23] := 'U';
       ELSIF "Control_DB".LCnv_Sys[1].Cnv_Level[1].Cnv2.Pallet_Type = 3 THEN
           "DB_Send_Data_To_Logistex".VTD_J1310_OUTFEED.Pallet_ID[23] := 'E';
       END_IF;

       // 2
       "Handshake_Outfeed_FC"(Auto_Mode := "Control_DB".LCnv_Sys[2].Cnv_Level[1].Cnv2.Mode = 3,
                              Ready_To_Send := "Control_DB".LCnv_Sys[2].Cnv_Level[1].Cnv2.Instruction.Outbound_Ready,
                              Conv_Occupied := "Control_DB".LCnv_Sys[2].Cnv_Level[1].Cnv2.Cnv_Occupied,
                              Transfer_In_Progress := "Control_DB".LCnv_Sys[2].Cnv_Level[1].Cnv2.Running,
                              DB_LGX_To_SM_Outfeed_Ready_To_Receive := "DB_Receive_Data_From_Logistex".J1320_Conv_Oufeed.LGXReadyToReceive,
                              Fault_Handshake => #Fault_Handshake_Outfeed_2,
                              DB_SM_To_LGX_Outfeed_Transfer_In_Progress => "DB_Send_Data_To_Logistex".VTD_J1320_OUTFEED.SPMTransferingInProgress,
                              DB_SM_To_LGX_Outfeed_Ocuppied => "DB_Send_Data_To_Logistex".VTD_J1320_OUTFEED.SPMTransferingOccupied,
                              DB_SM_To_LGX_Outfeed_Ready_To_Send => "DB_Send_Data_To_Logistex".VTD_J1320_OUTFEED.SPMReadyToSend);

       // Pallet tpe
       IF "Control_DB".LCnv_Sys[2].Cnv_Level[1].Cnv2.Pallet_Type = 1 THEN
           "DB_Send_Data_To_Logistex".VTD_J1320_OUTFEED.Pallet_ID[23] := 'U';
       ELSIF "Control_DB".LCnv_Sys[2].Cnv_Level[1].Cnv2.Pallet_Type = 3 THEN
           "DB_Send_Data_To_Logistex".VTD_J1320_OUTFEED.Pallet_ID[23] := 'E';
       END_IF;

       // 3
       "Handshake_Outfeed_FC"(Auto_Mode := "Control_DB".LCnv_Sys[3].Cnv_Level[1].Cnv2.Mode = 3,
                              Ready_To_Send := "Control_DB".LCnv_Sys[3].Cnv_Level[1].Cnv2.Instruction.Outbound_Ready,
                              Conv_Occupied := "Control_DB".LCnv_Sys[3].Cnv_Level[1].Cnv2.Cnv_Occupied,
                              Transfer_In_Progress := "Control_DB".LCnv_Sys[3].Cnv_Level[1].Cnv2.Running,
                              DB_LGX_To_SM_Outfeed_Ready_To_Receive := "DB_Receive_Data_From_Logistex".J1330_Conv_Oufeed.LGXReadyToReceive,
                              Fault_Handshake => #Fault_Handshake_Outfeed_3,
                              DB_SM_To_LGX_Outfeed_Transfer_In_Progress => "DB_Send_Data_To_Logistex".VTD_J1330_OUTFEED.SPMTransferingInProgress,
                              DB_SM_To_LGX_Outfeed_Ocuppied => "DB_Send_Data_To_Logistex".VTD_J1330_OUTFEED.SPMTransferingOccupied,
                              DB_SM_To_LGX_Outfeed_Ready_To_Send => "DB_Send_Data_To_Logistex".VTD_J1330_OUTFEED.SPMReadyToSend);

       // Pallet tpe
       IF "Control_DB".LCnv_Sys[3].Cnv_Level[1].Cnv2.Pallet_Type = 1 THEN
           "DB_Send_Data_To_Logistex".VTD_J1330_OUTFEED.Pallet_ID[23] := 'U';
       ELSIF "Control_DB".LCnv_Sys[3].Cnv_Level[1].Cnv2.Pallet_Type = 3 THEN
           "DB_Send_Data_To_Logistex".VTD_J1330_OUTFEED.Pallet_ID[23] := 'E';
       END_IF;
   END_REGION ;

   REGION STATUS
       REGION SEND
           "VTD_Status_Update_FC"(
                                  Infeed_Auto_Mode := "Control_DB".LCnv_Sys[1].Cnv_Level[1].Cnv1.Mode = 3,
                                  Infeed_Manual_Mode := "Control_DB".LCnv_Sys[1].Cnv_Level[1].Cnv1.Mode <> 3,
                                  Infeed_Maintenance := "Control_DB".VTD_Sys[1].Mode = 5,
                                  Infeed_Alarm := "Control_DB".LCnv_Sys[1].Cnv_Level[1].Cnv1.Error,
                                  Infeed_Ready := "Control_DB".LCnv_Sys[1].Cnv_Level[1].Cnv1.Instruction.Inbound_Ready,
                                  Outfeed_Auto_Mode := "Control_DB".LCnv_Sys[1].Cnv_Level[1].Cnv2.Mode = 3,
                                  Pallet_ID := "DB_Receive_Data_From_Logistex".J1310_Conv_Infeed.Pallet_ID,
                                  Pallet_ID_Received := "Control_DB".Pallet_ID_Received[1],
                                  SM_To_LGX_VTD_Status => "DB_Send_Data_To_Logistex".VTD_STATUS[1]
           );

           "VTD_Status_Update_FC"(
                                  Infeed_Auto_Mode := "Control_DB".LCnv_Sys[2].Cnv_Level[1].Cnv1.Mode = 3,
                                  Infeed_Manual_Mode := "Control_DB".LCnv_Sys[2].Cnv_Level[1].Cnv1.Mode <> 3,
                                  Infeed_Maintenance := "Control_DB".VTD_Sys[2].Mode = 5,
                                  Infeed_Alarm := "Control_DB".LCnv_Sys[2].Cnv_Level[1].Cnv1.Error,
                                  Infeed_Ready := "Control_DB".LCnv_Sys[2].Cnv_Level[1].Cnv1.Instruction.Inbound_Ready,
                                  Outfeed_Auto_Mode := "Control_DB".LCnv_Sys[2].Cnv_Level[1].Cnv2.Mode = 3,
                                  Pallet_ID := "DB_Receive_Data_From_Logistex".J1320_Conv_Infeed.Pallet_ID,
                                  Pallet_ID_Received := "Control_DB".Pallet_ID_Received[2],
                                  SM_To_LGX_VTD_Status => "DB_Send_Data_To_Logistex".VTD_STATUS[2]
           );

           "VTD_Status_Update_FC"(
                                  Infeed_Auto_Mode := "Control_DB".LCnv_Sys[3].Cnv_Level[1].Cnv1.Mode = 3,
                                  Infeed_Manual_Mode := "Control_DB".LCnv_Sys[3].Cnv_Level[1].Cnv1.Mode <> 3,
                                  Infeed_Maintenance := "Control_DB".VTD_Sys[3].Mode = 5,
                                  Infeed_Alarm := "Control_DB".LCnv_Sys[3].Cnv_Level[1].Cnv1.Error,
                                  Infeed_Ready := "Control_DB".LCnv_Sys[3].Cnv_Level[1].Cnv1.Instruction.Inbound_Ready,
                                  Outfeed_Auto_Mode := "Control_DB".LCnv_Sys[3].Cnv_Level[1].Cnv2.Mode = 3,
                                  Pallet_ID := "DB_Receive_Data_From_Logistex".J1330_Conv_Infeed.Pallet_ID,
                                  Pallet_ID_Received := "Control_DB".Pallet_ID_Received[3],
                                  SM_To_LGX_VTD_Status => "DB_Send_Data_To_Logistex".VTD_STATUS[3]
           );

           "DB_Send_Data_To_Logistex".PLC_STATUS.Hardbit := "Clock_1Hz";
           "DB_Send_Data_To_Logistex".PLC_STATUS."PLC_E-Stop" := "System_DB_1".Error AND "System_DB_2".Error AND "System_DB_3".Error;

           //Light guard and gate status
           "DB_Send_Data_To_Logistex".VTD_STATUS[4].%X0 := "Remote_Panel_DB_1".Light_Guards_CX101.Q;
           "DB_Send_Data_To_Logistex".VTD_STATUS[4].%X1 := "Remote_Panel_DB_2".Light_Guards_CX101.Q;
           "DB_Send_Data_To_Logistex".VTD_STATUS[4].%X2 := "Remote_Panel_DB_3".Light_Guards_CX101.Q;
           "DB_Send_Data_To_Logistex".VTD_STATUS[4].%X3 := "Remote_Panel_DB_1".Light_Guards_CX201.Q;
           "DB_Send_Data_To_Logistex".VTD_STATUS[4].%X4 := "Remote_Panel_DB_2".Light_Guards_CX201.Q;
           "DB_Send_Data_To_Logistex".VTD_STATUS[4].%X5 := "Remote_Panel_DB_3".Light_Guards_CX201.Q;

           //Gates
           "DB_Send_Data_To_Logistex".VTD_STATUS[5].%X0 := "Remote_Panel_DB_1".Gate_1_DB.Q;
           "DB_Send_Data_To_Logistex".VTD_STATUS[5].%X1 := "Remote_Panel_DB_1".Gate_2_DB.Q;
           "DB_Send_Data_To_Logistex".VTD_STATUS[5].%X2 := "Remote_Panel_DB_2".Gate_1_DB.Q;
           "DB_Send_Data_To_Logistex".VTD_STATUS[5].%X3 := "Remote_Panel_DB_2".Gate_2_DB.Q;
           "DB_Send_Data_To_Logistex".VTD_STATUS[5].%X4 := "Remote_Panel_DB_3".Gate_1_DB.Q;
           "DB_Send_Data_To_Logistex".VTD_STATUS[5].%X5 := "Remote_Panel_DB_3".Gate_2_DB.Q;

           //Requested Access
           "DB_Send_Data_To_Logistex".VTD_STATUS[6].%X0 := "GateAccess_Station_FB_DB_1".CurrentState <> #AUTO_RUNNING OR "GateAccess_Station_FB_DB_2".CurrentState <> #AUTO_RUNNING;
           "DB_Send_Data_To_Logistex".VTD_STATUS[6].%X1 := "GateAccess_Station_FB_DB_3".CurrentState <> #AUTO_RUNNING OR "GateAccess_Station_FB_DB_4".CurrentState <> #AUTO_RUNNING;
           "DB_Send_Data_To_Logistex".VTD_STATUS[6].%X2 := "GateAccess_Station_FB_DB_5".CurrentState <> #AUTO_RUNNING OR "GateAccess_Station_FB_DB_6".CurrentState <> #AUTO_RUNNING;

           //Speed conveyors 
           "DB_Send_Data_To_Logistex".CONV_SPEED.VTD_J1310_INF_SP := UINT_TO_INT("Settings_DB".LCnv_Sys[1].Cnv_Level[1].Cnv1.Full_Speed);
           "DB_Send_Data_To_Logistex".CONV_SPEED.VTD_J1310_OUF_SP := UINT_TO_INT("Settings_DB".LCnv_Sys[1].Cnv_Level[1].Cnv2.Full_Speed);
           "DB_Send_Data_To_Logistex".CONV_SPEED.VTD_J1320_INF_SP := UINT_TO_INT("Settings_DB".LCnv_Sys[2].Cnv_Level[1].Cnv1.Full_Speed);
           "DB_Send_Data_To_Logistex".CONV_SPEED.VTD_J1320_OUF_SP := UINT_TO_INT("Settings_DB".LCnv_Sys[2].Cnv_Level[1].Cnv2.Full_Speed);
           "DB_Send_Data_To_Logistex".CONV_SPEED.VTD_J1330_INF_SP_1 := UINT_TO_INT("Settings_DB".LCnv_Sys[3].Cnv_Level[1].Cnv1.Full_Speed);
           "DB_Send_Data_To_Logistex".CONV_SPEED.VTD_J1330_OUF_SP := UINT_TO_INT("Settings_DB".LCnv_Sys[3].Cnv_Level[1].Cnv2.Full_Speed);

       END_REGION

       REGION RECEIVE
           "LGX_ReadyToReceive_1" := "DB_Receive_Data_From_Logistex".J1310_Conv_Oufeed.LGXTransferingInProgress AND NOT "DB_Receive_Data_From_Logistex".CNV_STATUS[4].%X7; //Running and no error
           "LGX_ReadyToReceive_2" := "DB_Receive_Data_From_Logistex".J1320_Conv_Oufeed.LGXTransferingInProgress AND NOT "DB_Receive_Data_From_Logistex".CNV_STATUS[5].%X7;
           "LGX_ReadyToReceive_3" := "DB_Receive_Data_From_Logistex".J1330_Conv_Oufeed.LGXTransferingInProgress AND NOT "DB_Receive_Data_From_Logistex".CNV_STATUS[6].%X7;

           //Guaranteed Access 
           "LGX_Secure_Access_1" := "DB_Receive_Data_From_Logistex".CNV_STATUS[7].%X0;
           "LGX_Secure_Access_2" := "DB_Receive_Data_From_Logistex".CNV_STATUS[7].%X1;
           "LGX_Secure_Access_3" := "DB_Receive_Data_From_Logistex".CNV_STATUS[7].%X2;
       END_REGION
   END_REGION ;
END_FUNCTION

FUNCTION "FC_CLOCK" : DTL   // FC55, LAD
{ S7_Optimized_Access := 'TRUE' }
VERSION : 0.1
// stored: AutoNumber true, IsIECCheckEnabled false, SetENOAutomatically false, UDAEnableTagReadback false
   VAR_OUTPUT
      CurrentTime : String;
   END_VAR
   VAR_TEMP
      CurrentDTL : DTL;
      RetVal : Int;
      TempString : String;
      strYear : String;
      strMonth : String;
      strDay : String;
      strHour : String;
      strMinute : String;
      strSeconds : String;
   END_VAR
   VAR_TEMP   // added for the SCL form of the ladder/FBD networks
      _w1 : Bool;
      _w2 : Bool;
      _w3 : Bool;
      _w4 : Bool;
      _w5 : Bool;
   END_VAR
BEGIN

REGION Network 1: Read Current Local Time
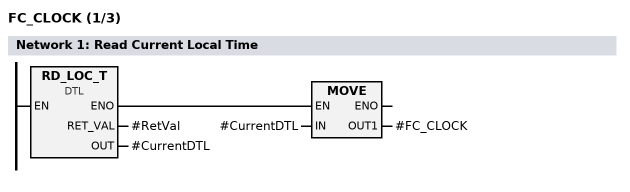
   RUNG wire#powerrail
      { S7_Templates := "date_type := DTL" } RD_LOC_T(RET_VAL => #RetVal, OUT => #CurrentDTL)
      Move(in := #CurrentDTL, out1 => #FC_CLOCK)
   END_RUNG
   // the same network as SCL:
   #RetVal := RD_LOC_T(OUT => #CurrentDTL, ENO => #_w1);
   IF #_w1 THEN #FC_CLOCK := #CurrentDTL; END_IF;
END_REGION

